(* IEC 61131-3 sources: Antarbhukti-LLM/DatasetCreation/SeedSTs/batch2_filtered_NETWORK, 29 files *)

(* ---- DLOG_FILE_TO_FTP.ST ---- *)
(*@PROPERTIES_EX@
TYPE: POU
LOCALE: 0
IEC_LANGUAGE: ST
PLC_TYPE: independent
PROC_TYPE: independent
GROUP: DATA_LOG
*)
(*@KEY@:DESCRIPTION*)
version 1.1		26. jul. 2011
programmer		ks
tested by		ks

DLOG_FILE_TO_FTP der Baustein kopiert bzw verschiebt die vom DLOG_STORE_FILE_CSV erzeugten Dateien auf einem FTP-Server

(*@KEY@:END_DESCRIPTION*)
FUNCTION_BLOCK DLOG_FILE_TO_FTP

(*Group:parameter*)

VAR_INPUT
	FTP_URL :	oscat_STRING250;
	FTP_ACTIV :	BOOL;
	FILE_DELETE :	BOOL;
	TIMEOUT :	TIME := T#30s;
	RETRY :	INT;
	RETRY_TIME :	TIME := T#30s;
	DNS_IP4 :	DWORD;
	PLC_IP4 :	DWORD;
END_VAR

VAR_OUTPUT
	DONE :	BOOL;
	BUSY :	BOOL;
	ERROR_C :	DWORD;
	ERROR_T :	BYTE;
END_VAR

VAR_IN_OUT
	X :	oscat_DLOG_DATA;
END_VAR

(*Group:lokal*)

VAR
	UCBD :	oscat_UNI_CIRCULAR_BUFFER_DATA;
	UCB :	UNI_CIRCULAR_BUFFER;
	FTP_CLIENT :	FTP_CLIENT;
	WT_1 :	TON;
	ftrig_old :	BOOL;
	filename :	STRING;
	step :	INT;
	ftp_busy :	BOOL;
	ftp_done :	BOOL;
	cnt :	INT;
END_VAR

(*Group:debug*)

VAR
	(*<LOG_MSG :	LOG_MSG;>*)
END_VAR

VAR_EXTERNAL
	(*<LOG_CL :	us_LOG_CONTROL;>*)(*Debug-Datenstruktur*)
END_VAR

VAR
	(*<_debug_enable :	BOOL := TRUE;>*)
END_VAR

(*@KEY@: WORKSHEET
NAME: DLOG_FILE_TO_FTP
IEC_LANGUAGE: ST
*)
(* neue Filenamen speichern *)
IF X.NEW_FILE_RTRIG AND ftrig_old = FALSE THEN
	UCBD.D_HEAD := WORD#1;
	UCBD.D_MODE := 1;
	UCBD.D_STRING := X.NEW_FILE;
	UCB(DATA:=UCBD); (* Daten eintragen *)
	UCBD := UCB.DATA;
END_IF;
ftrig_old := X.NEW_FILE_RTRIG;

CASE step OF

00:	IF UCBD.BUF_COUNT > 0 AND ftp_busy = FALSE THEN
		UCBD.D_MODE := 12; (* Daten lesen und löschen *)
		UCB(DATA:=UCBD);
		UCBD := UCB.DATA;
		filename := UCBD.D_STRING;
		cnt := 0;
		step := 10;
	END_IF;

10:	IF ftp_busy = FALSE THEN
		IF ftp_done THEN
			(*####################  DEBUG-MESSAGE  ###################################*)
			(*IF _debug_enable THEN
				LOG_CL.NEW_MSG := 'F_T_FTP: /FILE OK >~1<';
				LOG_CL.PRINTF[1] := filename;
				LOG_MSG();
			END_IF;*)
			(*########################################################################*)
			step := 0;
		ELSE
			step := 20; (* pause nach error *)
		END_IF;
	END_IF;

20:	IF WT_1.Q THEN (* Wartezeit *)
		cnt := cnt - 1;
		IF RETRY = 0 THEN (* FTP Transfer unbegrenzt wiederholen *)
			(*####################  DEBUG-MESSAGE  ###################################*)
			(*IF _debug_enable THEN
				LOG_CL.NEW_MSG := 'F_T_FTP: Auftrag unbegrenzt wiederholen /file: ~2';
				LOG_CL.PRINTF[2] := filename;
				LOG_MSG();
			END_IF;*)
			(*########################################################################*)
			step := 10; (* FTP Transfer wiederholen *)
		ELSIF cnt >= 0 THEN
			(*####################  DEBUG-MESSAGE  ###################################*)
			(*IF _debug_enable THEN
				LOG_CL.NEW_MSG := 'F_T_FTP: Auftrag wiederholen /cnt: ~1 /file: ~2';
				LOG_CL.PRINTF[1] := INT_TO_STRING(cnt,'%d');
				LOG_CL.PRINTF[2] := filename;
				LOG_MSG();
			END_IF;*)
			(*########################################################################*)
			step := 10; (* FTP Transfer wiederholen *)
		ELSE
			(*####################  DEBUG-MESSAGE  ###################################*)
			(*IF _debug_enable THEN
				LOG_CL.NEW_MSG := 'F_T_FTP: Auftrag verworfen /file: ~2';
				LOG_CL.PRINTF[2] := filename;
				LOG_MSG();
			END_IF;*)
			(*########################################################################*)
			step := 0; (* FTP Auftrag verwerfen *)
		END_IF;
	END_IF;

END_CASE;

BUSY := step = 10;
DONE := step = 0;
WT_1(IN:= step = 20, PT:= RETRY_TIME);

FTP_CLIENT(
	ACTIVATE:= BUSY,
	FILENAME:= filename,
	FTP_URL:= FTP_URL,
	FTP_DOWNLOAD:= FALSE,
	FTP_ACTIV:= FTP_ACTIV,
	FILE_DELETE:= FILE_DELETE,
	TIMEOUT:= TIMEOUT,
	DNS_IP4:= DNS_IP4,
	PLC_IP4:= PLC_IP4
	);
	ftp_done := FTP_CLIENT.DONE;
	ftp_busy := FTP_CLIENT.BUSY;
	ERROR_C := FTP_CLIENT.ERROR_C;
	ERROR_T := FTP_CLIENT.ERROR_T;

(* revision history
ks	01. jan. 2011	rev 1.0
	original version

ks	26. jul. 2011	rev 1.1
    codeoptimierung D_MODE 12

*)

(*@KEY@: END_WORKSHEET *)
END_FUNCTION_BLOCK

(* ---- DLOG_FILE_TO_SMTP.ST ---- *)
(*@PROPERTIES_EX@
TYPE: POU
LOCALE: 0
IEC_LANGUAGE: ST
PLC_TYPE: independent
PROC_TYPE: independent
GROUP: DATA_LOG
*)
(*@KEY@:DESCRIPTION*)
version 1.2		26. jul. 2011
programmer		ks
tested by		ks

DLOG_FILE_TO_SMTP der Baustein versendet die vom DLOG_STORE_FILE_CSV erzeugten Dateien als Email

(*@KEY@:END_DESCRIPTION*)
FUNCTION_BLOCK DLOG_FILE_TO_SMTP

(*Group:parameter*)

VAR_INPUT
	FILE_DELETE :	BOOL;
	TIMEOUT :	TIME := T#30s;
	DTI :	UDINT;
	DTI_OFFSET :	INT;
	RETRY :	INT;
	RETRY_TIME :	TIME := T#30s;
	DNS_IP4 :	DWORD;
END_VAR

VAR_OUTPUT
	DONE :	BOOL;
	BUSY :	BOOL;
	ERROR_C :	DWORD;
	ERROR_T :	BYTE;
END_VAR

VAR_IN_OUT
	SERVER :	STRING;
	MAILFROM :	STRING;
	MAILTO :	oscat_STRING250;
	SUBJECT :	STRING;
	BODY :	oscat_STRING250;
	X :	oscat_DLOG_DATA;
END_VAR

(*Group:lokal*)

VAR
	UCBD :	oscat_UNI_CIRCULAR_BUFFER_DATA;
	UCB :	UNI_CIRCULAR_BUFFER;
	SMTP_CLIENT :	SMTP_CLIENT;
	WT_1 :	TON;
	ftrig_old :	BOOL;
	files :	oscat_STRING250;
	step :	INT;
	smtp_busy :	BOOL;
	smtp_done :	BOOL;
	cnt :	INT;
END_VAR

(*Group:debug*)

VAR
	(*<LOG_MSG :	LOG_MSG;>*)
END_VAR

VAR_EXTERNAL
	(*<LOG_CL :	us_LOG_CONTROL;>*)(*Debug-Datenstruktur*)
END_VAR

VAR
	(*<_debug_enable :	BOOL := TRUE;>*)
END_VAR

(*@KEY@: WORKSHEET
NAME: DLOG_FILE_TO_SMTP
IEC_LANGUAGE: ST
*)
(* neue Filenamen speichern *)
IF X.NEW_FILE_RTRIG AND ftrig_old = FALSE THEN
	UCBD.D_HEAD := WORD#1;
	UCBD.D_MODE := 1;
	UCBD.D_STRING := X.NEW_FILE;
	UCB(DATA:=UCBD); (* Daten eintragen *)
	UCBD := UCB.DATA;
END_IF;
ftrig_old := X.NEW_FILE_RTRIG;

CASE step OF

00:	IF UCBD.BUF_COUNT > 0 AND smtp_busy = FALSE THEN
		UCBD.D_MODE := 12; (* Daten lesen und löschen *)
		UCB(DATA:=UCBD);
		UCBD := UCB.DATA;
		files := UCBD.D_STRING;
		IF FILE_DELETE THEN
			files := CONCAT(files,';#DEL#');
		END_IF;
		cnt := 0;
		step := 10;
	END_IF;

10:	IF smtp_busy = FALSE THEN
		IF smtp_done THEN
			(*####################  DEBUG-MESSAGE  ###################################*)
			(*IF _debug_enable THEN
				LOG_CL.NEW_MSG := 'F_T_SMTP: /FILE OK >~1<';
				LOG_CL.PRINTF[1] := files;
				LOG_MSG();
			END_IF;*)
			(*########################################################################*)
			step := 0;
		ELSE
			step := 20; (* pause nach error *)
		END_IF;
	END_IF;

20:	IF WT_1.Q THEN (* Wartezeit *)
		cnt := cnt - 1;
		IF RETRY = 0 THEN (* Transfer unbegrenzt wiederholen *)
			(*####################  DEBUG-MESSAGE  ###################################*)
			(*IF _debug_enable THEN
				LOG_CL.NEW_MSG := 'F_T_SMTP: Auftrag unbegrenzt wiederholen /file: ~2';
				LOG_CL.PRINTF[2] := files;
				LOG_MSG();
			END_IF;*)
			(*########################################################################*)
			step := 10; (* Transfer wiederholen *)
		ELSIF cnt >= 0 THEN
			(*####################  DEBUG-MESSAGE  ###################################*)
			(*IF _debug_enable THEN
				LOG_CL.NEW_MSG := 'F_T_SMTP: Auftrag wiederholen /cnt: ~1 /file: ~2';
				LOG_CL.PRINTF[1] := INT_TO_STRING(cnt,'%d');
				LOG_CL.PRINTF[2] := files;
				LOG_MSG();
			END_IF;*)
			(*########################################################################*)
			step := 10; (* Transfer wiederholen *)
		ELSE
			(*####################  DEBUG-MESSAGE  ###################################*)
			(*IF _debug_enable THEN
				LOG_CL.NEW_MSG := 'F_T_SMTP: Auftrag verworfen /file: ~2';
				LOG_CL.PRINTF[2] := files;
				LOG_MSG();
			END_IF;*)
			(*########################################################################*)
			step := 0; (* Auftrag verwerfen *)
		END_IF;
	END_IF;

END_CASE;

BUSY := step = 10;
DONE := step = 0;
WT_1(IN:= step = 20, PT:= RETRY_TIME);

SMTP_CLIENT(
	ACTIVATE:= BUSY,
	TIMEOUT:= TIMEOUT,
	DTI:= DTI,
	DTI_OFFSET:= DTI_OFFSET,
	DNS_IP4:= DNS_IP4,
	SERVER:= SERVER,
	MAILFROM:= MAILFROM,
	MAILTO:= MAILTO,
	SUBJECT:= SUBJECT,
	BODY:= BODY,
	FILES:= FILES
	);
	SERVER:= SMTP_CLIENT.SERVER;
	MAILFROM:= SMTP_CLIENT.MAILFROM;
	MAILTO:= SMTP_CLIENT.MAILTO;
	SUBJECT:= SMTP_CLIENT.SUBJECT;
	BODY:= SMTP_CLIENT.BODY;
	FILES:= SMTP_CLIENT.FILES;
	smtp_done := SMTP_CLIENT.DONE;
	smtp_busy := SMTP_CLIENT.BUSY;
	ERROR_C := SMTP_CLIENT.ERROR_C;
	ERROR_T := SMTP_CLIENT.ERROR_T;

(* revision history

ks	01. jan. 2011	rev 1.0
	original version

ks	28. apr. 2011	rev 1.1
	stringfehler bei option 'file_delete'

ks	26. jul. 2011	rev 1.2
    codeoptimierung D_MODE 12
*)

(*@KEY@: END_WORKSHEET *)
END_FUNCTION_BLOCK

(* ---- DLOG_STORE_FILE_CSV.ST ---- *)
(*@PROPERTIES_EX@
TYPE: POU
LOCALE: 0
IEC_LANGUAGE: ST
PLC_TYPE: independent
PROC_TYPE: independent
GROUP: DATA_LOG
*)
(*@KEY@:DESCRIPTION*)
version 1.2		25. jul. 2011
programmer		ks
tested by		ks

DLOG_STORE_FILE_CSV der Baustein schreibt die DLOG Parameter in einen lokale Datei im CSV-Format

(*@KEY@:END_DESCRIPTION*)
FUNCTION_BLOCK DLOG_STORE_FILE_CSV

(*Group:Default*)

VAR_INPUT
	ENABLE :	BOOL;
	TRIG_M :	BOOL;
	TRIG_T :	UDINT;
	FILENAME :	STRING;
	DTI :	UDINT;
	SEP :	BYTE;
END_VAR

VAR_OUTPUT
	ERROR_C :	DWORD;
	ERROR_T :	BYTE;
END_VAR

VAR_IN_OUT
	X :	oscat_DLOG_DATA;
END_VAR

VAR
	FS :	FILE_SERVER;
	FSD :	oscat_FILE_SERVER_DATA;
	PT :	oscat_NETWORK_BUFFER;
	UCB :	UNI_CIRCULAR_BUFFER;
	ra :	BOOL;
	trig_m_last :	BOOL;
	dti_last :	UDINT := udint#4294967295;(*DT#2070-02-06-06:28:15*)
	enable_last :	BOOL;
	fn_last :	STRING;
	fn :	STRING;
	init :	BOOL;
	step :	INT;
	idx :	INT;
	log_stop :	BOOL;
	buf_totalsize :	INT := 4096;
	DT_TO_STRF :	DT_TO_STRF;
	_STRING_TO_BUFFER :	_STRING_TO_BUFFER_NW;
	n :	USINT;
END_VAR

(*@KEY@: WORKSHEET
NAME: DLOG_STORE_FILE_CSV
IEC_LANGUAGE: ST
*)
X.DTI := DTI; (* Datum / Zeit eintragen *)
IF DTI <> dti_last THEN
	X.CLOCK_TRIG := TRUE;
	dti_last := DTI;
	X.STORE_TYPE := BYTE#2;
ELSE
	X.CLOCK_TRIG := FALSE;
END_IF;

IF X.ADD_HEADER = FALSE THEN (* wenn add-header und add-data gleichzeitig ansteht, dann add-data einen zyklus länger anstehen lassen *)
	X.ADD_DATA := FALSE;
END_IF;
X.ADD_HEADER := FALSE;

IF ENABLE THEN
	IF X.CLOCK_TRIG THEN
		DT_TO_STRF(DTI:=DTI,MS:=0,FMT:=FILENAME,LANG:=0); (* automatische Dateinamen generierung *)
		fn := DT_TO_STRF.DT_TO_STRF;
		IF TRIG_T > UDINT#0 THEN (* automatischer Trigger *)
			ra := DTI MOD TRIG_T = UDINT#0;
		END_IF;
	ELSE
		ra := FALSE;
	END_IF;
	IF (TRIG_M AND NOT trig_m_last) OR ra THEN (* manueller oder automatischer Trigger *)
		X.ADD_DATA := TRUE; (* Daten loggen *)
	END_IF;
	IF NOT init THEN
		init := TRUE;
		X.ADD_HEADER := TRUE; (* Spaltenüberschriften übernehmen *)
	END_IF;
END_IF;

IF (NOT ENABLE AND enable_last) OR (NE_STRING(fn,fn_last) AND step > 0) THEN (* Neg. Flanke ENABLE - Log Stop *)
	fn_last := fn;
	X.UCB.D_HEAD := WORD#16#FF00;
	X.UCB.D_MODE := 1;
	UCB(DATA:=X.UCB); (* Element schreiben *)
	X.UCB := UCB.DATA;
	X.ADD_HEADER := TRUE; (* Spaltenüberschriften übernehmen *)
END_IF;

CASE step OF

00:	IF ENABLE THEN
		fn_last := fn;
		FSD.FILENAME := fn; (* Dateiname *)
		FSD.OFFSET := UDINT#0; (* Start bei Dateianfang *)
		FSD.AUTO_CLOSE := T#0s; (* Auto-Close *)
		step := 20;
	END_IF;

20:	IF X.UCB.BUF_COUNT > 0 THEN (* Einträge vorhanden *)
		X.UCB.D_MODE := 10;
		UCB(DATA:=X.UCB); (* Element lesen , aber noch nicht entfernen *)
		X.UCB := UCB.DATA;
		IF X.UCB.D_HEAD = WORD#16#FF00 THEN (* LOG_STOP Command *)
			X.UCB.D_MODE := 11;
			UCB(DATA:=X.UCB); (* Element entfernen *)
			X.UCB := UCB.DATA;
			log_stop := TRUE;
			step := 40; (* Daten schreiben *)
		ELSIF idx + LEN(X.UCB.D_STRING) + 2 < buf_totalsize THEN (* Platz für Element vorhanden ? *)
			X.UCB.D_MODE := 11;
			UCB(DATA:=X.UCB); (* Element entfernen *)
			X.UCB := UCB.DATA;
			_STRING_TO_BUFFER(STR:=X.UCB.D_STRING, POS:=idx, PT:=PT.BUFFER, SIZE:=INT_TO_UINT(buf_totalsize));
			PT.BUFFER:=_STRING_TO_BUFFER.PT;
			idx := idx + LEN(X.UCB.D_STRING);
			n := n + USINT#1;
			IF n = X.ID_MAX THEN (* letztes Element einer Zeile *)
				n := USINT#0;
				PT.BUFFER[idx] := BYTE#16#0D;
				idx := idx + 1;
				PT.BUFFER[idx] := BYTE#16#0A;
			ELSE
				PT.BUFFER[idx] := SEP;
			END_IF;
			idx := idx + 1;
		ELSE
			step := 40; (* Daten schreiben *)
		END_IF;
	END_IF;

40:	IF idx > 0 THEN (* Daten schreiben *)
		FSD.MODE := BYTE#3; (* create + write *)
		PT.SIZE := INT_TO_UINT(idx); (* Datenlänge eintragen *)
		idx := 0;
	END_IF;
	step := 60;

60:	IF FSD.MODE = BYTE#0 THEN
		IF log_stop THEN
			log_stop := FALSE;
			FSD.MODE := BYTE#5; (* Datei schliessen *)
			X.NEW_FILE := FSD.FILENAME;
			X.NEW_FILE_RTRIG := FALSE;
			step := 80;
		ELSE
			step := 20;
		END_IF;
	END_IF;

80:	IF FSD.MODE = BYTE#0 THEN (* Datei schliessen beendet *)
		X.NEW_FILE_RTRIG := TRUE;
		step := 0;
	END_IF;

END_CASE;

trig_m_last := TRIG_M;
enable_last := ENABLE;

FS(FSD:=FSD,PT:=PT); (* FILE_SERVER *)
FSD := FS.FSD;
PT  := FS.PT;

ERROR_C := BYTE_TO_DWORD(FSD.ERROR);
ERROR_T := SEL(FSD.ERROR > BYTE#0,BYTE#0,BYTE#1);

(* revision history
ks	01. jan. 2011	rev 1.0
	original version

ks	13. may. 2011	rev 1.1
	ADD_DATA_REQ, ERROR_T, ERROR_C hinzugefügt

ks	25. jul. 2011	rev 1.2
	HEAD informationen geändert, neuer Spaltenzähler

*)

(*@KEY@: END_WORKSHEET *)
END_FUNCTION_BLOCK

(* ---- DLOG_STORE_FILE_HTML.ST ---- *)
(*@PROPERTIES_EX@
TYPE: POU
LOCALE: 0
IEC_LANGUAGE: ST
PLC_TYPE: independent
PROC_TYPE: independent
GROUP: DATA_LOG
*)
(*@KEY@:DESCRIPTION*)

(*@KEY@:END_DESCRIPTION*)
FUNCTION_BLOCK DLOG_STORE_FILE_HTML

(*Group:Default*)

VAR_INPUT
	ENABLE :	BOOL;
	TRIG_M :	BOOL;
	TRIG_T :	UDINT;
	FILENAME :	STRING;
	DTI :	UDINT;
	HTML_CAPTION :	STRING;
	HTML_TABLE :	STRING;
	HTML_TR_HEAD :	STRING;
	HTML_TR_EVEN :	STRING;
	HTML_TR_ODD :	STRING;
END_VAR

VAR_OUTPUT
	ERROR_C :	DWORD;
	ERROR_T :	BYTE;
END_VAR

VAR_IN_OUT
	X :	oscat_DLOG_DATA;
END_VAR

VAR
	FS :	FILE_SERVER;
	FSD :	oscat_FILE_SERVER_DATA;
	PT :	oscat_NETWORK_BUFFER;
	UCB :	UNI_CIRCULAR_BUFFER;
	ra :	BOOL;
	trig_m_last :	BOOL;
	dti_last :	UDINT := udint#4294967295;(*DT#2070-02-06-06:28:15*)
	enable_last :	BOOL;
	fn_last :	STRING;
	str :	oscat_STRING250;
	fn :	STRING;
	init :	BOOL;
	step :	INT;
	idx :	INT;
	log_state :	USINT;
	color :	BOOL;
	head :	BOOL;
	n :	USINT;
	buf_totalsize :	INT := 4096;
	DT_TO_STRF :	DT_TO_STRF;
	_STRING_TO_BUFFER :	_STRING_TO_BUFFER_NW;
END_VAR

(*@KEY@: WORKSHEET
NAME: DLOG_STORE_FILE_HTML
IEC_LANGUAGE: ST
*)
X.DTI := DTI; (* Datum / Zeit eintragen *)
IF DTI <> dti_last THEN
	X.CLOCK_TRIG := TRUE;
	dti_last := DTI;
	X.STORE_TYPE := BYTE#4;
ELSE
	X.CLOCK_TRIG := FALSE;
END_IF;

IF X.ADD_HEADER = FALSE THEN (* wenn add-header und add-data gleichzeitig ansteht, dann add-data einen zyklus länger anstehen lassen *)
	X.ADD_DATA := FALSE;
END_IF;
X.ADD_HEADER := FALSE;

IF ENABLE THEN
	IF X.CLOCK_TRIG THEN
		DT_TO_STRF(DTI:=DTI,MS:=0,FMT:=FILENAME,LANG:=0); (* automatische Dateinamen generierung *)
		fn := DT_TO_STRF.DT_TO_STRF;
		IF TRIG_T > UDINT#0 THEN (* automatischer Trigger *)
			ra := DTI MOD TRIG_T = UDINT#0;
		END_IF;
	ELSE
		ra := FALSE;
	END_IF;
	IF (TRIG_M AND NOT trig_m_last) OR ra OR X.ADD_DATA_REQ THEN (* manueller, automatischer oder externer Trigger *)
		X.ADD_DATA := TRUE; (* Daten loggen *)
	END_IF;
	IF NOT init THEN
		init := TRUE;
		X.ADD_HEADER := TRUE; (* Spaltenüberschriften übernehmen *)
	END_IF;
END_IF;
X.ADD_DATA_REQ := FALSE; (* externe Anforderung rücksetzen *)

IF (NOT ENABLE AND enable_last) OR (NE_STRING(fn,fn_last) AND step > 0) THEN (* Neg. Flanke ENABLE - Log Stop *)
	fn_last := fn;
	X.UCB.D_HEAD := WORD#16#FF00;
	X.UCB.D_MODE := 1;
	UCB(DATA:=X.UCB); (* Element schreiben *)
	X.UCB := UCB.DATA;
	X.ADD_HEADER := TRUE; (* Spaltenüberschriften übernehmen *)
END_IF;

CASE step OF

00:	IF ENABLE THEN
		color := FALSE;
		head := FALSE;
		fn_last := fn;
		FSD.FILENAME := fn; (* Dateiname *)
		FSD.OFFSET := UDINT#0; (* Start bei Dateianfang *)
		FSD.AUTO_CLOSE := T#0s; (* Auto-Close *)
		step := 10;
	END_IF;

10:	(* Headerdaten schreiben *)
	str := CONCAT('<html><body><table ',HTML_TABLE);
	str := CONCAT(str,'><caption>');
	str := CONCAT(str,HTML_CAPTION);
	str := CONCAT(str,'</caption>');

	_STRING_TO_BUFFER(STR:=str, POS:=idx, PT:=PT.BUFFER, SIZE:=INT_TO_UINT(buf_totalsize));
	PT.BUFFER:=_STRING_TO_BUFFER.PT;
	idx := idx + LEN(str);
	step := 20;

20:	IF log_state = USINT#254 THEN
		log_state := USINT#255;
		str := '</table></body></html>';
		_STRING_TO_BUFFER(STR:=str, POS:=idx, PT:=PT.BUFFER, SIZE:=INT_TO_UINT(buf_totalsize));
		PT.BUFFER:=_STRING_TO_BUFFER.PT;
		idx := idx + LEN(str);
		step := 40; (* Daten schreiben *)

	ELSIF X.UCB.BUF_COUNT > 0 THEN (* Einträge vorhanden *)
		X.UCB.D_MODE := 10;
		UCB(DATA:=X.UCB); (* Element lesen , aber noch nicht entfernen *)
		X.UCB := UCB.DATA;

		IF X.UCB.D_HEAD = WORD#16#FF00 THEN (* LOG_STOP Command *)
			X.UCB.D_MODE := 11;
			UCB(DATA:=X.UCB); (* Element entfernen *)
			X.UCB := UCB.DATA;
			log_state := USINT#254;

		ELSIF idx + LEN(X.UCB.D_STRING) + 120 < buf_totalsize THEN (* Platz für Element vorhanden ? *)
			X.UCB.D_MODE := 11;
			UCB(DATA:=X.UCB); (* Element entfernen *)
			X.UCB := UCB.DATA;

			IF log_state = USINT#0 THEN
				str := '<TR ';
				IF NOT head THEN
					str := CONCAT(str,HTML_TR_HEAD);
					head := TRUE;
				ELSIF color THEN
					str := CONCAT(str,HTML_TR_EVEN);
				ELSE
					str := CONCAT(str,HTML_TR_ODD);
				END_IF;
				str := CONCAT(str,'><TD>');
			ELSE
				str := '<TD>';
			END_IF;
			_STRING_TO_BUFFER(STR:=str, POS:=idx, PT:=PT.BUFFER, SIZE:=INT_TO_UINT(buf_totalsize));
			PT.BUFFER:=_STRING_TO_BUFFER.PT;
			idx := idx + LEN(str);
			log_state := log_state + USINT#1;

			_STRING_TO_BUFFER(STR:=X.UCB.D_STRING, POS:=idx, PT:=PT.BUFFER, SIZE:=INT_TO_UINT(buf_totalsize));
			PT.BUFFER:=_STRING_TO_BUFFER.PT;
			idx := idx + LEN(X.UCB.D_STRING);
			n := n + USINT#1;
			IF n = X.ID_MAX THEN
				n := USINT#0;
				str := '</TD></TR>';
				color := NOT color;
				log_state := USINT#0;
			ELSE
				str := '</TD>';
			END_IF;
			_STRING_TO_BUFFER(STR:=str, POS:=idx, PT:=PT.BUFFER, SIZE:=INT_TO_UINT(buf_totalsize));
			PT.BUFFER:=_STRING_TO_BUFFER.PT;
			idx := idx + LEN(str);
		END_IF;
		step := 40; (* Daten schreiben *)
	END_IF;

40:	IF idx > 0 THEN (* Daten schreiben *)
		FSD.MODE := BYTE#3; (* create + write *)
		PT.SIZE := INT_TO_UINT(idx); (* Datenlänge eintragen *)
		idx := 0;
	END_IF;
	step := 60;

60:	IF FSD.MODE = BYTE#0 THEN
		IF log_state = USINT#255 THEN
			log_state := USINT#0;
			FSD.MODE := BYTE#5; (* Datei schliessen *)
			X.NEW_FILE := FSD.FILENAME;
			X.NEW_FILE_RTRIG := FALSE;
			step := 80;
		ELSE
			step := 20;
		END_IF;
	END_IF;

80:	IF FSD.MODE = BYTE#0 THEN (* Datei schliessen beendet *)
		X.NEW_FILE_RTRIG := TRUE;
		step := 0;
	END_IF;

END_CASE;

trig_m_last := TRIG_M;
enable_last := ENABLE;

FS(FSD:=FSD,PT:=PT); (* FILE_SERVER *)
FSD := FS.FSD;
PT  := FS.PT;

ERROR_C := BYTE_TO_DWORD(FSD.ERROR);
ERROR_T := SEL(FSD.ERROR > BYTE#0,BYTE#0,BYTE#1);

(* revision history
ks	25. july. 2011	rev 1.0
	original version

*)

(*@KEY@: END_WORKSHEET *)
END_FUNCTION_BLOCK

(* ---- DLOG_STORE_FILE_XML.ST ---- *)
(*@PROPERTIES_EX@
TYPE: POU
LOCALE: 0
IEC_LANGUAGE: ST
PLC_TYPE: independent
PROC_TYPE: independent
GROUP: DATA_LOG
*)
(*@KEY@:DESCRIPTION*)
version 1.0		25. july. 2011
programmer		ks
tested by		ks

DLOG_STORE_FILE_XML schreibt die DLOG Parameter in einen lokale Datei im XML-Format

(*@KEY@:END_DESCRIPTION*)
FUNCTION_BLOCK DLOG_STORE_FILE_XML

(*Group:Default*)

VAR_INPUT
	ENABLE :	BOOL;
	TRIG_M :	BOOL;
	TRIG_T :	UDINT;
	FILENAME :	STRING;
	DTI :	UDINT;
END_VAR

VAR_OUTPUT
	ERROR_C :	DWORD;
	ERROR_T :	BYTE;
END_VAR

VAR_IN_OUT
	X :	oscat_DLOG_DATA;
END_VAR

VAR
	FS :	FILE_SERVER;
	FSD :	oscat_FILE_SERVER_DATA;
	PT :	oscat_NETWORK_BUFFER;
	UCB :	UNI_CIRCULAR_BUFFER;
	ra :	BOOL;
	trig_m_last :	BOOL;
	dti_last :	UDINT := udint#4294967295;(*DT#2070-02-06-06:28:15*)
	enable_last :	BOOL;
	fn_last :	STRING;
	str :	oscat_STRING250;
	fn :	STRING;
	init :	BOOL;
	step :	INT;
	idx :	INT;
	log_state :	USINT;
	n :	USINT;
	buf_totalsize :	INT := 4096;
	DT_TO_STRF :	DT_TO_STRF;
	_STRING_TO_BUFFER :	_STRING_TO_BUFFER_NW;
END_VAR

(*@KEY@: WORKSHEET
NAME: DLOG_STORE_FILE_XML
IEC_LANGUAGE: ST
*)
X.DTI := DTI; (* Datum / Zeit eintragen *)
IF DTI <> dti_last THEN
	X.CLOCK_TRIG := TRUE;
	dti_last := DTI;
	X.STORE_TYPE := BYTE#3;
ELSE
	X.CLOCK_TRIG := FALSE;
END_IF;

IF X.ADD_HEADER = FALSE THEN (* wenn add-header und add-data gleichzeitig ansteht, dann add-data einen zyklus länger anstehen lassen *)
	X.ADD_DATA := FALSE;
END_IF;
X.ADD_HEADER := FALSE;

IF ENABLE THEN
	IF X.CLOCK_TRIG THEN
		DT_TO_STRF(DTI:=DTI,MS:=0,FMT:=FILENAME,LANG:=0); (* automatische Dateinamen generierung *)
		fn := DT_TO_STRF.DT_TO_STRF;
		IF TRIG_T > UDINT#0 THEN (* automatischer Trigger *)
			ra := DTI MOD TRIG_T = UDINT#0;
		END_IF;
	ELSE
		ra := FALSE;
	END_IF;
	IF (TRIG_M AND NOT trig_m_last) OR ra OR X.ADD_DATA_REQ THEN (* manueller, automatischer oder externer Trigger *)
		X.ADD_DATA := TRUE; (* Daten loggen *)
	END_IF;
	IF NOT init THEN
		init := TRUE;
		X.ADD_HEADER := TRUE; (* Spaltenüberschriften übernehmen *)
	END_IF;
END_IF;
X.ADD_DATA_REQ := FALSE; (* externe Anforderung rücksetzen *)

IF (NOT ENABLE AND enable_last) OR (NE_STRING(fn,fn_last) AND step > 0) THEN (* Neg. Flanke ENABLE - Log Stop *)
	fn_last := fn;
	X.UCB.D_HEAD := WORD#16#FF00;
	X.UCB.D_MODE := 1;
	UCB(DATA:=X.UCB); (* Element schreiben *)
	X.UCB := UCB.DATA;
	X.ADD_HEADER := TRUE; (* Spaltenüberschriften übernehmen *)
END_IF;

CASE step OF

00:	IF ENABLE THEN
		fn_last := fn;
		FSD.FILENAME := fn; (* Dateiname *)
		FSD.OFFSET := UDINT#0; (* Start bei Dateianfang *)
		FSD.AUTO_CLOSE := T#0s; (* Auto-Close *)
		step := 10;
	END_IF;

10:	(* Headerdaten schreiben *)
	str := '<?xml version="1.0" encoding="UTF-8"?><table>';
	_STRING_TO_BUFFER(STR:=str, POS:=idx, PT:=PT.BUFFER, SIZE:=INT_TO_UINT(buf_totalsize));
	PT.BUFFER:=_STRING_TO_BUFFER.PT;
	idx := idx + LEN(str);
	step := 20;

20:	IF log_state = USINT#254 THEN
		log_state := USINT#255;
		str := '</table>';
		_STRING_TO_BUFFER(STR:=str, POS:=idx, PT:=PT.BUFFER, SIZE:=INT_TO_UINT(buf_totalsize));
		PT.BUFFER:=_STRING_TO_BUFFER.PT;
		idx := idx + LEN(str);
		step := 40; (* Daten schreiben *)

	ELSIF X.UCB.BUF_COUNT > 0 THEN (* Einträge vorhanden *)
		X.UCB.D_MODE := 10;
		UCB(DATA:=X.UCB); (* Element lesen , aber noch nicht entfernen *)
		X.UCB := UCB.DATA;

		IF X.UCB.D_HEAD = WORD#16#FF00 THEN (* LOG_STOP Command *)
			X.UCB.D_MODE := 11;
			UCB(DATA:=X.UCB); (* Element entfernen *)
			X.UCB := UCB.DATA;
			log_state := USINT#254;

		ELSIF idx + LEN(X.UCB.D_STRING) + 120 < buf_totalsize THEN (* Platz für Element vorhanden ? *)
			X.UCB.D_MODE := 11;
			UCB(DATA:=X.UCB); (* Element entfernen *)
			X.UCB := UCB.DATA;

			IF log_state = USINT#0 THEN
				str := '<row><entry>';
			ELSE
				str := '<entry>';
			END_IF;

			_STRING_TO_BUFFER(STR:=str, POS:=idx, PT:=PT.BUFFER, SIZE:=INT_TO_UINT(buf_totalsize));
			PT.BUFFER:=_STRING_TO_BUFFER.PT;
			idx := idx + LEN(str);
			log_state := log_state + USINT#1;

			_STRING_TO_BUFFER(STR:=X.UCB.D_STRING, POS:=idx, PT:=PT.BUFFER, SIZE:=INT_TO_UINT(buf_totalsize));
			PT.BUFFER:=_STRING_TO_BUFFER.PT;
			idx := idx + LEN(X.UCB.D_STRING);

			n := n + USINT#1;
			IF n = X.ID_MAX THEN
				n := USINT#0;
				str := '</entry></row>';
				log_state := USINT#0;
			ELSE
				str := '</entry>';
			END_IF;
			_STRING_TO_BUFFER(STR:=str, POS:=idx, PT:=PT.BUFFER, SIZE:=INT_TO_UINT(buf_totalsize));
			PT.BUFFER:=_STRING_TO_BUFFER.PT;
			idx := idx + LEN(str);
		END_IF;
		step := 40; (* Daten schreiben *)
	END_IF;

40:	IF idx > 0 THEN (* Daten schreiben *)
		FSD.MODE := BYTE#3; (* create + write *)
		PT.SIZE := INT_TO_UINT(idx); (* Datenlänge eintragen *)
		idx := 0;
	END_IF;
	step := 60;

60:	IF FSD.MODE = BYTE#0 THEN
		IF log_state = USINT#255 THEN
			log_state := USINT#0;
			FSD.MODE := BYTE#5; (* Datei schliessen *)
			X.NEW_FILE := FSD.FILENAME;
			X.NEW_FILE_RTRIG := FALSE;
			step := 80;
		ELSE
			step := 20;
		END_IF;
	END_IF;

80:	IF FSD.MODE = BYTE#0 THEN (* Datei schliessen beendet *)
		X.NEW_FILE_RTRIG := TRUE;
		step := 0;
	END_IF;

END_CASE;

trig_m_last := TRIG_M;
enable_last := ENABLE;

FS(FSD:=FSD,PT:=PT); (* FILE_SERVER *)
FSD := FS.FSD;
PT  := FS.PT;

ERROR_C := BYTE_TO_DWORD(FSD.ERROR);
ERROR_T := SEL(FSD.ERROR > BYTE#0,BYTE#0,BYTE#1);

(* revision history
ks	25. july. 2011	rev 1.0
	original version

*)
(*@KEY@: END_WORKSHEET *)
END_FUNCTION_BLOCK

(* ---- DLOG_STORE_RRD.ST ---- *)
(*@PROPERTIES_EX@
TYPE: POU
LOCALE: 0
IEC_LANGUAGE: ST
PLC_TYPE: independent
PROC_TYPE: independent
GROUP: DATA_LOG
*)
(*@KEY@:DESCRIPTION*)
version 1.2		26. jul. 2011
programmer		ks
tested by		ks

DLOG_STORE_RRD der Baustein übergibt die DLOG Parameter an einen RoundRobinDatabase-Server

(*@KEY@:END_DESCRIPTION*)
FUNCTION_BLOCK DLOG_STORE_RRD

(*Group:Default*)

VAR_INPUT
	ENABLE :	BOOL;
	TRIG_M :	BOOL;
	TRIG_T :	UDINT;
	URL :	oscat_STRING250;
	DTI :	UDINT;
	SEP :	BYTE;
	DNS_IP4 :	DWORD;
	TIMEOUT :	TIME;
END_VAR

VAR_OUTPUT
	ERROR_C :	DWORD;
	ERROR_T :	BYTE;
END_VAR

VAR_IN_OUT
	X :	oscat_DLOG_DATA;
END_VAR

VAR
	UCB :	UNI_CIRCULAR_BUFFER;
	IP_C :	oscat_IP_C;
	S_BUF :	oscat_NETWORK_BUFFER;
	R_BUF :	oscat_NETWORK_BUFFER;
	URL_DATA :	oscat_url;
	DNS_CLIENT :	DNS_CLIENT;
	HTTP_GET :	HTTP_GET;
	IPC :	IP_CONTROL;
	ra :	BOOL;
	trig_m_last :	BOOL;
	dti_last :	UDINT := udint#4294967295;(*DT#2070-02-06-06:28:15*)
	step :	INT;
	sep_char :	oscat_STRING1;
	STRING_TO_URL :	STRING_TO_URL;
	CHR_TO_STRING :	CHR_TO_STRING;
	n :	INT;
END_VAR

(*@KEY@: WORKSHEET
NAME: DLOG_STORE_RRD
IEC_LANGUAGE: ST
*)
X.DTI := DTI; (* Datum / Zeit eintragen *)
IF DTI <> dti_last THEN
	X.CLOCK_TRIG := TRUE;
	dti_last := DTI;
	X.STORE_TYPE := BYTE#1;
ELSE
	X.CLOCK_TRIG := FALSE;
END_IF;

X.ADD_DATA := FALSE;

IF ENABLE THEN
	IF X.CLOCK_TRIG THEN
		IF TRIG_T > UDINT#0 THEN (* automatischer Trigger *)
			ra := DTI MOD TRIG_T = UDINT#0;
		END_IF;
	ELSE
		ra := FALSE;
	END_IF;
	IF (TRIG_M AND NOT trig_m_last) OR ra OR X.ADD_DATA_REQ THEN (* manueller, automatischer oder externer Trigger *)
		X.ADD_DATA := TRUE; (* Daten loggen *)
	END_IF;
END_IF;
X.ADD_DATA_REQ := FALSE; (* externe Anforderung rücksetzen *)

CASE step OF

00:	IF ENABLE THEN
		STRING_TO_URL(STR:=URL,DEFAULT_PROTOCOL:='',DEFAULT_PATH:=''); (* URL zerlegen *)
		URL_DATA:=STRING_TO_URL.STRING_TO_URL;
		CHR_TO_STRING(C:=SEP);
		sep_char:=CHR_TO_STRING.CHR_TO_STRING;
		ERROR_T := BYTE#0;
		ERROR_C := DWORD#0;
		step := 20;
	END_IF;

20:	IF X.UCB.BUF_COUNT >= USINT_TO_INT(X.ID_MAX) THEN (* Einträge vorhanden *)
		n := 1;
		WHILE n <= USINT_TO_INT(X.ID_MAX) DO
			X.UCB.D_MODE := 12; (* Element lesen und löschen *)
			UCB(DATA:=X.UCB);
			X.UCB := UCB.DATA;
			IF n < USINT_TO_INT(X.ID_MAX) THEN (* Trennzeichen hinzufügen *)
				X.UCB.D_STRING := CONCAT(X.UCB.D_STRING,sep_char);
			END_IF;
			IF LEN(X.UCB.D_STRING) + LEN(URL_DATA.QUERY) <= 250 THEN
				URL_DATA.QUERY := CONCAT(URL_DATA.QUERY,X.UCB.D_STRING); (* Query mit LOG-Daten ergänzen *)
				step :=40;
			ELSE
				ERROR_T := BYTE#4; (* LOG-Daten können nicht in URL gepackt werden *)
				ERROR_C := DWORD#1;
				step := 0;
			END_IF;
			n := n + 1;
		END_WHILE;;
	END_IF;

40:	IF DNS_CLIENT.DONE THEN
		step := 60;
	ELSIF (DNS_CLIENT.ERROR > DWORD#0) THEN
		ERROR_C := DNS_CLIENT.ERROR; (* Fehlerbehandlung *)
		ERROR_T := BYTE#1;
		step := 100;
	END_IF;

60:	IF HTTP_GET.DONE THEN
		n := UINT_TO_INT(HTTP_GET.BODY_START);
		IF R_BUF.BUFFER[n] <> BYTE#48 THEN (* ASCII '0' *)
			ERROR_C := DWORD#1;
			ERROR_T := BYTE#3;
		END_IF;
		step := 100;

	ELSIF HTTP_GET.ERROR > DWORD#0 THEN (* Fehlerbehandlung *)
		ERROR_C := HTTP_GET.ERROR;
		ERROR_T := BYTE#2;
		step := 100;
	END_IF;

100:	IF (NOT HTTP_GET.DONE) THEN (* UNLOCK HTTP DATA *)
		step := SEL(ERROR_T = BYTE#0, 120,0);
	END_IF;

120:	IF NOT ENABLE THEN
		X.UCB.D_MODE := 99;
		UCB(DATA:=X.UCB); (* Buffer löschen *)
		X.UCB := UCB.DATA;
		step := 0;
	END_IF;

END_CASE;

HTTP_GET(IP_C:=IP_C,S_BUF:=S_BUF,R_BUF:=R_BUF,IP4:=DNS_CLIENT.IP4,GET:=step=60,MODE:=BYTE#2,UNLOCK_BUF:=step=100,URL_DATA:=URL_DATA); (* HTTP_GET *)
IP_C     := HTTP_GET.IP_C;
S_BUF    := HTTP_GET.S_BUF;
R_BUF    := HTTP_GET.R_BUF;
URL_DATA := HTTP_GET.URL_DATA;

DNS_CLIENT(IP_C:=IP_C, S_BUF:=S_BUF, R_BUF:=R_BUF, DOMAIN:=URL_DATA.DOMAIN, IP4_DNS:= DNS_IP4, ACTIVATE:=step=40); (* DNS-Client *)
IP_C  := DNS_CLIENT.IP_C;
S_BUF := DNS_CLIENT.S_BUF;
R_BUF := DNS_CLIENT.R_BUF;

IPC(IP:= DWORD#0, PORT:= WORD#0 , TIME_OUT:= TIMEOUT, IP_C:= IP_C, S_BUF:= S_BUF, R_BUF:= R_BUF); (* IP_CONTROL *)
IP_C  := IPC.IP_C;
S_BUF := IPC.S_BUF;
R_BUF := IPC.R_BUF;

trig_m_last := TRIG_M;

(* revision history
ks	01. jan. 2011	rev 1.0
	original version

ks	13. may. 2011	rev 1.1
	ADD_DATA_REQ hinzugefügt

ks	26. july. 2011	rev 1.2
	code optimierung D_MODE 12 und bessere fehlerauswertung
*)

(*@KEY@: END_WORKSHEET *)
END_FUNCTION_BLOCK

(* ---- DNS_CLIENT.ST ---- *)
(*@PROPERTIES_EX@
TYPE: POU
LOCALE: 0
IEC_LANGUAGE: ST
PLC_TYPE: independent
PROC_TYPE: independent
GROUP: NETWORK
*)
(*@KEY@:DESCRIPTION*)

version 1.3		26. jul. 2011
programmer 		ks
tested by		ks

DNS_CLIENT führt eine Domain-Name Abfrage bei einen DNS-Server durch
(*@KEY@:END_DESCRIPTION*)
FUNCTION_BLOCK DNS_CLIENT

(*Group:log*)

VAR
	(*<LOG_MSG :	LOG_MSG;>*)
	(*<_debug_enable :	BOOL := FALSE;>*)
END_VAR

VAR_EXTERNAL
	(*<LOG_CL :	us_LOG_CONTROL;>*)
END_VAR

(*Group:lokal*)

VAR
	IP4_DECODE :	IP4_DECODE;
	IP_FIFO :	IP_FIFO;
	CODE :	CODE;
	ip_state :	BYTE;
	ip_id :	BYTE;
	i :	INT;
	i1 :	INT;
	i2 :	INT;
	i3 :	INT;
	state :	INT;
	domain_copy :	STRING;
	activate_last :	BOOL;
	url_length :	INT;
	char :	BYTE;
	char_count :	INT;
	tid :	BYTE;
	anc :	INT;
	x :	BYTE;
	rr_stop :	BOOL;
	ttl_last :	DWORD;
	ttl_tmp :	DWORD;
	z :	INT;
END_VAR

(*Group:Default*)

VAR_IN_OUT
	IP_C :	oscat_IP_C;(*IP_Control Verwaltungsstruktur*)
	S_BUF :	oscat_NETWORK_BUFFER;
	R_BUF :	oscat_NETWORK_BUFFER;
END_VAR

VAR_INPUT
	ACTIVATE :	BOOL;
	DOMAIN :	STRING;
	IP4_DNS :	DWORD;
END_VAR

VAR_OUTPUT
	IP4 :	DWORD;
	DONE :	BOOL;
	ERROR :	DWORD;
END_VAR

(*@KEY@: WORKSHEET
NAME: DNS_CLIENT
IEC_LANGUAGE: ST
*)
(* Domain Name System (query) *)

CASE state OF

00:	IF ACTIVATE AND NOT activate_last THEN (* auf positive Flanke GET warten *)
		DONE := FALSE;
		ERROR := DWORD#0;
		state := 5;
	END_IF;

05: (* prüfe ob domain schon eine IP4-Adresse ist *)
    IP4_DECODE(str:=DOMAIN);
    IP4 := IP4_DECODE.IP4_DECODE; (* IP4 Adresse direkt weitergeben *)
	IF IP4 > DWORD#00 THEN
		DONE := TRUE;
		state := 0;
        (*####################  DEBUG-MESSAGE  ###################################*)
        (*IF _debug_enable THEN
            LOG_CL.NEW_MSG := 'DNS: S05 IP4 ~1';
            LOG_CL.PRINTF[1]  := DOMAIN;
            LOG_MSG();
        END_IF;*)
        (*########################################################################*)
	ELSE
		ip_state := BYTE#1;
		ttl_last := DWORD#0;
		domain_copy := DOMAIN; (* DOMAIN String sichern *)
		state := 10;
        (*####################  DEBUG-MESSAGE  ###################################*)
        (*IF _debug_enable THEN
            LOG_CL.NEW_MSG := 'DNS: S05 START';
            LOG_MSG();
        END_IF;*)
        (*########################################################################*)
	END_IF;

10:	IF ip_state = BYTE#3 THEN (* Bei IP_Control anmelden *)
		url_length := LEN(domain_copy);
		char_count := 17 + url_length; (* sendebuffer initialisieren *)
		FOR i := 0 TO char_count DO
			S_BUF.BUFFER[i] := BYTE#00;
		END_FOR;
		tid := UINT_TO_BYTE(BYTE_TO_UINT(tid) + UINT#1);
		S_BUF.BUFFER[01] := tid; (* Transaction ID lowbyte *)
		S_BUF.BUFFER[02] := BYTE#16#01; (* Flags: highbyte *)
		S_BUF.BUFFER[05] := BYTE#16#01; (* Questions: lowbyte *)
		i := url_length + 12; (* den servernamen von hinten nach vorne bearbeiten *)
		char_count := 0;
		WHILE i > 12 DO
			CODE(STR:=domain_copy,POS:=i - 12);
			char := CODE.CODE;
			IF char = BYTE#46 THEN (* prüfe auf haupt/sub domänen namens-teiler "." *)
				S_BUF.BUFFER[i] := INT_TO_BYTE(char_count); (* anstelle des teilers "." wird die länge des erkannten haupt/sub domänennames eingetragen *)
				char_count := 0;
			ELSE
				S_BUF.BUFFER[i] := char; (* char in buffer eintragen *)
				char_count := char_count + 1; (* anzahl char zählen *)
			END_IF;
			i := i - 1;
		END_WHILE;
		S_BUF.BUFFER[i] := INT_TO_BYTE(char_count); (* längenangabe des ganz linken (ersten) domänennamens eintragen *)
		i := url_length + 15; (* position hinter dem servernamen *)
		S_BUF.BUFFER[i] := BYTE#01; (* Type: A Hostaddress lowbyte *)
		i := i + 2;
		S_BUF.BUFFER[i] := BYTE#01; (* Class: IN lowbyte *)
		i := i + 1;
		(* IP Datenverkehr einrichten *)
		IP_C.C_PORT := WORD#53; (* Portnummer eintragen *)
		IP_C.C_IP := IP4_DNS; (* IP eintragen *)
		IP_C.C_MODE := BYTE#1; (* Mode: UDP+AKTIV+PORT+IP *)
		IP_C.C_ENABLE := TRUE; (* Verbindungsaufbau freigeben *)
		IP_C.TIME_RESET := TRUE; (* Zeitueberwachung rücksetzen *)
		IP_C.R_OBSERVE  := TRUE; (* Datenempfang ueberwachen *)
		S_BUF.SIZE := INT_TO_UINT(i); (* sendelänge eintragen *)
		R_BUF.SIZE := UINT#0; (* Empfangslänge rücksetzen *)
		state := 30;

        (*####################  DEBUG-MESSAGE  ###################################*)
        (*IF _debug_enable THEN
            LOG_CL.NEW_MSG := 'DNS: S10 SEND';
            LOG_MSG();
        END_IF;*)
        (*########################################################################*)
	END_IF;

30:	IF IP_C.ERROR <> DWORD#00 THEN
		ERROR := IP_C.ERROR;
		state := 99;
        (*####################  DEBUG-MESSAGE  ###################################*)
        (*IF _debug_enable THEN
            LOG_CL.NEW_MSG := 'DNS: S30 ERROR ~1';
            LOG_CL.PRINTF[1]  := DWORD_TO_STRING(ERROR,'%08X');
            LOG_MSG();
        END_IF;*)
        (*########################################################################*)

	ELSIF (S_BUF.SIZE = UINT#0) AND (tid = R_BUF.BUFFER[1]) AND (R_BUF.SIZE >= INT_TO_UINT(34 + url_length)) THEN	(* prüfe ob antwort telegramm die richtige Transaction-ID und mindestlänge hat *)
		ERROR := BYTE_TO_DWORD(R_BUF.BUFFER[3] AND BYTE#2#0000_1111); (* prüfe Return code der Flags. 4 bits *)
		IF ERROR = DWORD#00 THEN
			anc := _BYTE_TO_INT(R_BUF.BUFFER[7]); (* Anzahl der Answer-RR *)
			IP_C.R_OBSERVE := FALSE; (* Datenempfang ueberwachen *)
			state := 40;
		ELSE
			state := 99;
		END_IF;
	END_IF;

40:	IF anc > 0 THEN
		anc := anc - 1;
		z := UINT_TO_INT(R_BUF.SIZE);
		WHILE i < z DO
			x := R_BUF.BUFFER[i];
			IF rr_stop = FALSE THEN
				IF x > BYTE#63 THEN (* zeiger auf namen *)
					i := i + 1;
					rr_stop := TRUE;
				ELSIF x= BYTE#0 THEN (* namens ende *)
					rr_stop := TRUE;
				ELSE
					i := i + _BYTE_TO_INT(x); (* namen *)
				END_IF;
				i := i + 1;
			ELSE
				rr_stop := FALSE;
				i1 := i + 1;
				i3 := i + 3;
				IF R_BUF.BUFFER[i1] = BYTE#1 AND R_BUF.BUFFER[i3] = BYTE#1 THEN (* Type A / Class IN *)
					i := i + 4;
					i1 := i + 1;
					i2 := i + 2;
					i3 := i + 3;
					ttl_tmp := DWORD_OF_BYTE(R_BUF.BUFFER[i],R_BUF.BUFFER[i1],R_BUF.BUFFER[i2],R_BUF.BUFFER[i3]); (* Time to live *)
					i := i + 6;
					IF ttl_tmp >= ttl_last THEN (* TTL ist länger *)
						ttl_last := ttl_tmp;
						i1 := i + 1;
						i2 := i + 2;
						i3 := i + 3;
						IP4 := DWORD_OF_BYTE(R_BUF.BUFFER[i],R_BUF.BUFFER[i1],R_BUF.BUFFER[i2],R_BUF.BUFFER[i3]); (* IP-Adresse *)
					END_IF;
					i := i + 4;
				ELSE
					i := i + 9;
					i := i + _BYTE_TO_INT(R_BUF.BUFFER[i]) + 1; (* offset zu nächsten Block *)
				END_IF;
				EXIT;
			END_IF;
		END_WHILE;
	ELSE
		IF IP4 > DWORD#0 THEN (* gültige RR mit IP gefunden *)
			DONE := TRUE;
            (*####################  DEBUG-MESSAGE  ###################################*)
            (*IF _debug_enable THEN
                LOG_CL.NEW_MSG       := 'DNS: S40 OK';
                LOG_MSG();
            END_IF;*)
            (*########################################################################*)
		ELSE
			ERROR := DWORD#255; (* Daten fehlerhaft - keine IP-Adresse gefunden *)
		END_IF;
		state := 99;
	END_IF;

99:	R_BUF.SIZE := UINT#0; (* Empfangslänge rücksetzen *)
	ip_state := BYTE#4; (* Abmelden *)
	state := 00;

END_CASE;

activate_last := ACTIVATE; (* letzten Status sichern zur Flankenerkennung *)

IP_FIFO(FIFO:=IP_C.FIFO,STATE:=ip_state,ID:=ip_id); (* IP_FIFO *)
IP_C.FIFO:=IP_FIFO.FIFO;
ip_state := IP_FIFO.STATE;
ip_id:=IP_FIFO.ID;

(* revision history

ks	18. oct. 2008	rev 1.0
	original version

ks	20. oct. 2009	rev 1.1
	unbenutzten code entfernt, all buffer base 0

ks	20. dec. 2010	rev 1.2
	parsing nach rfc1305

ks	26. jul. 2011	rev 1.3
	verbesserte ip-auswertung, neue fehlermeldung
*)

(*----------------------------------------------------------------------------------------------------------------*)
(* Flags: 0x0100 (Standard query)                                                                                            *)
(* 0... .... .... .... = Response: Message is a query                                                                   *)
(* .000 0... ....  = Opcode: Standard query (0)                                                                          *)
(* .... ..0. .... .... = Truncated: Message is not truncated                                                          *)
(* .... ...1 .... .... = Recursion desired: Do query recursively                                                    *)
(* .... .... .0.. .... = Z: reserved (0)                                                                                                  *)
(* .... .... ...0 .... = Non-authenticated data OK: Non-authenticated data is unacceptable *)
(*-----------------------------------------------------------------------------------------------------------------*)

(*      0  1  2  3  4  5  6  7  8  9  0  1  2  3  4  5  *)
(*    +--+--+--+--+--+--+--+--+--+--+--+--+--+--+--+--+ *)
(*    |                      ID                       | idx: 0/1   *)
(*    +--+--+--+--+--+--+--+--+--+--+--+--+--+--+--+--+ *)
(*    |QR|   Opcode  |AA|TC|RD|RA|   Z    |   RCODE   | idx: 2/3   *)
(*    +--+--+--+--+--+--+--+--+--+--+--+--+--+--+--+--+ *)
(*    |                    QDCOUNT                    | idx: 4/5   *)
(*    +--+--+--+--+--+--+--+--+--+--+--+--+--+--+--+--+ *)
(*    |                    ANCOUNT                    | idx: 6/7   *)
(*    +--+--+--+--+--+--+--+--+--+--+--+--+--+--+--+--+ *)
(*    |                    NSCOUNT                    | idx: 8/9   *)
(*    +--+--+--+--+--+--+--+--+--+--+--+--+--+--+--+--+ *)
(*    |                    ARCOUNT                    | idx: 10/11 *)
(*    +--+--+--+--+--+--+--+--+--+--+--+--+--+--+--+--+ *)

(*
Errorcodes  Description	References
000	No error. 		 	The request completed successfully.
001	Format error. 		The name server was unable to interpret the query.
002	Server failure.  	The name server was unable to process this query due to a problem with the name server.
003	Name Error. 	 	Meaningful only for responses from an authoritative name server, this code signifies that the domain name referenced in the query does not exist.
004	Not Implemented. 	The name server does not support the requested kind of query.
005	Refused. 			The name server refuses to perform the specified operation for policy reasons.
  						 For example, a name server may not wish to provide the information to the particular requester, or a name server may not wish to perform a particular operation (e.g., zone transfer) for particular data.
006	YXDomain.			Name Exists when it should not.
007	YXRRSet. RR			Set Exists when it should not.
008	NXRRSet. RR			Set that should exist does not.
009	NotAuth.			Server Not Authoritative for zone.
010	NotZone,			Name not contained in zone.
255	Timeout				No Response

beispiel einer DNS Request von google.at
ein request mit 3 Answer-Blocks

Domain Name System (response)
[Request In: 3]
[Time: 0.027533000 seconds]
Transaction ID: 0x5e1a
Flags: 0x8180 (Standard query response, No error)
1... .... .... .... = Response: Message is a response
.000 0... .... .... = Opcode: Standard query (0)
.... .0.. .... .... = Authoritative: Server is not an authority for domain
.... ..0. .... .... = Truncated: Message is not truncated
.... ...1 .... .... = Recursion desired: Do query recursively
.... .... 1... .... = Recursion available: Server can do recursive queries
.... .... .0.. .... = Z: reserved (0)
.... .... ..0. .... = Answer authenticated: Answer/authority portion was not authenticated
.... .... .... 0000 = Reply code: No error (0)
Questions: 1
Answer RRs: 3
Authority RRs: 0
Additional RRs: 0

Queries
google.at: type A, class IN
Name: google.at
Type: A (Host address)
Class: IN (0x0001)

Answers
google.at: type A, class IN, addr 72.14.221.104
Name: google.at
Type: A (Host address)
Class: IN (0x0001)
Time to live: 19 minutes, 9 seconds
Data length: 4
Addr: 72.14.221.104

google.at: type A, class IN, addr 66.249.93.104
Name: google.at
Type: A (Host address)
Class: IN (0x0001)
Time to live: 19 minutes, 9 seconds
Data length: 4
Addr: 66.249.93.104

google.at: type A, class IN, addr 216.239.59.104
Name: google.at
Type: A (Host address)
Class: IN (0x0001)
Time to live: 19 minutes, 9 seconds
Data length: 4
Addr: 216.239.59.104
*)

(*@KEY@: END_WORKSHEET *)
END_FUNCTION_BLOCK

(* ---- DNS_REV_CLIENT.ST ---- *)
(*@PROPERTIES_EX@
TYPE: POU
LOCALE: 0
IEC_LANGUAGE: ST
PLC_TYPE: independent
PROC_TYPE: independent
GROUP: NETWORK
*)
(*@KEY@:DESCRIPTION*)
version 1.0	28. dec. 2009
programmer 	ks
tested BY	ks

DNS_REV_CLIENT führt eine Reverse-Domain-Name Abfrage durch, und ermittelt aus einer IP-Adresse den zugehörigen Domain-Namen.

(*@KEY@:END_DESCRIPTION*)
FUNCTION_BLOCK DNS_REV_CLIENT

(*Group:Default*)

VAR_IN_OUT
	IP_C :	oscat_IP_C;(*IP_Control Verwaltungsstruktur*)
	S_BUF :	oscat_NETWORK_BUFFER;
	R_BUF :	oscat_NETWORK_BUFFER;
END_VAR

VAR_INPUT
	ACTIVATE :	BOOL;
	IP4 :	DWORD;
	IP4_DNS :	DWORD;
END_VAR

VAR_OUTPUT
	DOMAIN :	STRING;
	DONE :	BOOL;
	ERROR :	DWORD;
END_VAR

VAR
	IP_FIFO :	IP_FIFO;
	ip_state :	BYTE;
	ip_id :	BYTE;
	state :	INT;
	ip4_copy :	DWORD;
	d :	oscat_STRING27;
	activate_last :	BOOL;
	i :	INT;
	dl :	INT;
	p1 :	INT;
	char :	BYTE;
	char_count :	INT;
	tid :	BYTE;
	BUFFER_TO_STRING :	BUFFER_TO_STRING_NW;
	CODE :	CODE;
END_VAR

(*@KEY@: WORKSHEET
NAME: DNS_REV_CLIENT
IEC_LANGUAGE: ST
*)
(* Domain Name System (query) *)

CASE state OF
00: (* auf positive Flanke GET warten *)
	IF ACTIVATE AND NOT activate_last THEN
		ERROR := DWORD#0;
		ip4_copy := ip4; (* IP4 sichern *)
		ip_state := BYTE#1;
		DOMAIN := '';
		DONE := FALSE;

		d := '';
		FOR i := 1 TO 4 DO
			d := CONCAT(d,BYTE_TO_STRING(DWORD_TO_BYTE(IP4),'%u'));
			d := CONCAT(d,'.');
			IP4 := ROR(IP4,8);
		END_FOR;
		d := CONCAT(d,'in-addr.arpa');
		state := 10;
	END_IF;

10: (* Bei IP_Control anmelden *)
	IF ip_state = BYTE#3 THEN
		dl := LEN(d);

		(* sendebuffer initialisieren *)
		char_count := 17 + dl;
		FOR i := 0 TO char_count DO
			S_BUF.BUFFER[i] := BYTE#00;
		END_FOR;

		tid := UINT_TO_BYTE(BYTE_TO_UINT(tid) + UINT#1);
		S_BUF.BUFFER[01] := tid; (* Transaction ID lowbyte *)
		S_BUF.BUFFER[02] := BYTE#16#01; (* Flags: highbyte *)
		S_BUF.BUFFER[05] := BYTE#16#01; (* Questions: lowbyte *)

		(* den servernamen von hinten nach vorne bearbeiten *)
		i := dl + 12;
		char_count := 0;

		WHILE i > 12 DO
			CODE(STR:=d,POS:=i - 12);
			char:=CODE.CODE;

			(* prüfe auf haupt/sub domänen namens-teiler "." *)
			IF char = BYTE#46 THEN
				(* anstelle des teilers "." wird die länge des erkannten haupt/sub domänennames eingetragen *)
				S_BUF.BUFFER[i] := INT_TO_BYTE(char_count);
				char_count := 0;
			ELSE
				S_BUF.BUFFER[i] := char; (* char in buffer eintragen *)
				char_count := char_count + 1; (* anzahl char zählen *)
			END_IF;
			i := i - 1;
		END_WHILE;

		S_BUF.BUFFER[i] := INT_TO_BYTE(char_count); (* längenangabe des ganz linken (ersten) domänennamens eintragen *)
		i := dl + 15; (* position hinter dem servernamen *)
		S_BUF.BUFFER[i] := BYTE#12; (* Type: PTR (Domain name pointer) lowbyte *)
		i := i + 2;
		S_BUF.BUFFER[i] := BYTE#01; (* Class: IN lowbyte *)
		i := i + 1;

		(* IP Datenverkehr einrichten *)
		IP_C.C_PORT := WORD#53; (* Portnummer eintragen *)
		IP_C.C_IP := IP4_DNS; (* IP eintragen *)
		IP_C.C_MODE := BYTE#1; (* Mode: UDP+AKTIV+PORT+IP *)
		IP_C.C_ENABLE := TRUE; (* Verbindungsaufbau freigeben *)
		IP_C.TIME_RESET := TRUE; (* Zeitueberwachung rücksetzen *)
		IP_C.R_OBSERVE  := TRUE; (* Datenempfang ueberwachen *)
		S_BUF.SIZE := INT_TO_UINT(i); (* sendelänge eintragen *)
		R_BUF.SIZE := UINT#0; (* Empfangslänge rücksetzen *)
		state := 30;
	END_IF;

30:
	IF IP_C.ERROR <> DWORD#00 THEN
		ERROR := IP_C.ERROR;
	(* prüfe ob antwort telegramm die richtige Transaction-ID und mindestlänge hat *)
	ELSIF (S_BUF.SIZE = UINT#0) AND (tid = R_BUF.BUFFER[1]) AND (R_BUF.SIZE >= INT_TO_UINT(i+12)) THEN

		(* prüfe Return code der Flags. 4 bits *)
		ERROR := BYTE_TO_DWORD(R_BUF.BUFFER[3] AND BYTE#2#0000_1111);

		IF ERROR = DWORD#00 THEN

			i := UINT_TO_INT(R_BUF.SIZE) - 2;
			WHILE R_BUF.BUFFER[i] > BYTE#0 DO
				IF i = 0 THEN EXIT; END_IF;
				i := i - 1;
			END_WHILE;

			i := i + 2;
			p1 := i + 1;
			WHILE i < UINT_TO_INT(R_BUF.SIZE) DO
				dl := _BYTE_TO_INT(R_BUF.BUFFER[i]);
				IF dl > 0 THEN
					R_BUF.BUFFER[i] := BYTE#46;
					i := i + dl + 1;
				ELSE

					BUFFER_TO_STRING(PT:=R_BUF.BUFFER,SIZE:=UINT#4096,START:=INT_TO_UINT(p1),STOP:=INT_TO_UINT(i-1));
					R_BUF.BUFFER:=BUFFER_TO_STRING.PT;
					DOMAIN:=BUFFER_TO_STRING.BUFFER_TO_STRING;
					EXIT;
				END_IF;
			END_WHILE;
			state := 0;
			DONE := TRUE;
		END_IF;
	END_IF;

	IF ERROR <> DWORD#0 THEN
		state := 0;
	END_IF;

	IF state = 0 THEN
		IP_C.R_OBSERVE := FALSE; (* Datenempfang ueberwachen *)
		ip_state := BYTE#4; (* Abmelden *)
	END_IF;

END_CASE;

activate_last := ACTIVATE; (* letzten Status sichern zur Flankenerkennung *)

(* IP_FIFO *)
IP_FIFO(FIFO:=IP_C.FIFO,STATE:=ip_state,ID:=ip_id);
IP_C.FIFO:=IP_FIFO.FIFO;
ip_state:=IP_FIFO.STATE;
ip_id:=IP_FIFO.ID;

(* revision history

ks	28. dec. 2009	rev 1.0
	original version

*)

(*----------------------------------------------------------------------------------------------------------------*)
(* Flags: 0x0100 (Standard query)                                                                                            *)
(* 0... .... .... .... = Response: Message is a query                                                                   *)
(* .000 0... ....  = Opcode: Standard query (0)                                                                          *)
(* .... ..0. .... .... = Truncated: Message is not truncated                                                          *)
(* .... ...1 .... .... = Recursion desired: Do query recursively                                                    *)
(* .... .... .0.. .... = Z: reserved (0)                                                                                                  *)
(* .... .... ...0 .... = Non-authenticated data OK: Non-authenticated data is unacceptable *)
(*-----------------------------------------------------------------------------------------------------------------*)

(*
Errorcodes  Description	References
000	No error. 		 	The request completed successfully.
001	Format error. 		The name server was unable to interpret the query.
002	Server failure.  	The name server was unable to process this query due to a problem with the name server.
003	Name Error. 	 	Meaningful only for responses from an authoritative name server, this code signifies that the domain name referenced in the query does not exist.
004	Not Implemented. 	The name server does not support the requested kind of query.
005	Refused. 			The name server refuses to perform the specified operation for policy reasons.
  						 For example, a name server may not wish to provide the information to the particular requester, or a name server may not wish to perform a particular operation (e.g., zone transfer) for particular data.
006	YXDomain.			Name Exists when it should not.
007	YXRRSet. RR			Set Exists when it should not.
008	NXRRSet. RR			Set that should exist does not.
009	NotAuth.			Server Not Authoritative for zone.
010	NotZone,			Name not contained in zone.
255	Timeout				No Response
*)

(*@KEY@: END_WORKSHEET *)
END_FUNCTION_BLOCK

(* ---- FILE_BLOCK.ST ---- *)
(*@PROPERTIES_EX@
TYPE: POU
LOCALE: 0
IEC_LANGUAGE: ST
PLC_TYPE: independent
PROC_TYPE: independent
GROUP: FILE
*)
(*@KEY@:DESCRIPTION*)
version 1.0		23. sep. 2010
programmer 		ks
tested by		ks

FILE_BLOCK liefert das angeforderte Byte einer Datei durch einlesen von möglichst grossen Datenblöcken

(*@KEY@:END_DESCRIPTION*)
FUNCTION_BLOCK FILE_BLOCK

(*Group:parameter*)

VAR_IN_OUT
	MODE :	BYTE;
	FILENAME :	STRING;
	FSD :	oscat_FILE_SERVER_DATA;
	PT :	oscat_NETWORK_BUFFER;
END_VAR

VAR_INPUT
	POS :	UDINT;
END_VAR

VAR_OUTPUT
	ERROR :	BYTE;
	DATA :	BYTE;
END_VAR

(*Group:log*)

VAR
	(*<LOG_MSG :	LOG_MSG;>*)
	(*<_debug_enable :	BOOL := TRUE;>*)
END_VAR

VAR_EXTERNAL
	(*<LOG_CL :	us_LOG_CONTROL;>*)
END_VAR

(*Group:var*)

VAR
	step :	INT;
	i :	INT;
	data_start :	UDINT;
	data_stop :	UDINT;
END_VAR

(*@KEY@: WORKSHEET
NAME: FILE_BLOCK
IEC_LANGUAGE: ST
*)
CASE step OF
0:	IF MODE > BYTE#0 THEN
		ERROR := BYTE#0;
		IF FSD.FILE_OPEN AND (FSD.FILE_SIZE = UDINT#0 OR POS >= FSD.FILE_SIZE) THEN
			ERROR := BYTE#255;
			MODE := BYTE#0;
		ELSIF POS < data_start OR POS > data_stop OR NOT FSD.FILE_OPEN THEN (* Daten lesen notwendig *)
			FSD.FILENAME := FILENAME;
			FSD.MODE := BYTE#1; (* open + read *)
			FSD.OFFSET := POS;
			PT.SIZE := UINT#65535; (* maximale anzahl lesen *);
			data_start := UDINT#0;
			data_stop := UDINT#0;
			step := 10;
		ELSE (* Daten sind im Buffer vorhanden *)
			i := UDINT_TO_INT(POS - data_start); (* index berechnen *)
			DATA := PT.BUFFER[i];
			MODE := BYTE#0;
			(* ---------------------- Debug-Message ----------------------------*)
			(*IF _debug_enable THEN
				LOG_CL.NEW_MSG := 'FB: Pos: ~1 Byte: ~2 >~3<';
				LOG_CL.PRINTF[1] := UDINT_TO_STRING(POS,'%03u');
				LOG_CL.PRINTF[2] := BYTE_TO_STRING(DATA,'%03u');
				LOG_CL.PRINTF[3] := BYTE_TO_STRING(DATA,'%c');
				LOG_MSG();
			END_IF;*)
			(* -----------------------------------------------------------------*)
		END_IF;
	END_IF;

10:	IF FSD.MODE = BYTE#0 THEN (* Befehl beendet *)
		IF FSD.ERROR > BYTE#0 THEN
			ERROR := FSD.ERROR; (* Fehler ausgeben *)
			MODE := BYTE#0;
		ELSE
			data_start := POS;
			data_stop := POS + UINT_TO_UDINT(PT.SIZE) - UDINT#1;
		END_IF;
		step := 0;
	END_IF;
END_CASE;

(* revision history
ks	23. sep. 2010	rev 1.0
	original version
*)

(*@KEY@: END_WORKSHEET *)
END_FUNCTION_BLOCK

(* ---- FILE_SERVER.ST ---- *)
(*@PROPERTIES_EX@
TYPE: POU
LOCALE: 0
IEC_LANGUAGE: ST
PLC_TYPE: independent
PROC_TYPE: independent
GROUP: HARDWARE
*)
(*@KEY@:DESCRIPTION*)
version 1.0		23. sep. 2010
programmer 		ks
tested by		ks

FILE_SERVER ermöglicht den Zugriff auf Dateien mittels Plattform-Neutraler Schnittstelle

Befehle:
1 = File_Open_Exist + File_Read
2 = File_Open_Exist + File_Write
3 = File_Open_New   + File_Write
4 = File_Remove
5 = File_Close

- Action -
1 = file_open   (open)
2 = file_close  (close)
3 = file_read   (read)
4 = file_write  (write)
5 = file_seek   (setpos)
6 = file_tell   (getpos)
7 = file_remove (delete)

---- fehlermeldungen----

000 (00) kein Fehler

002 (02) file_open - Die maximale Anzahl von Dateien ist bereits geöffnet.
004 (04) file_open - Die Datei ist bereits geöffnet.
005 (05) file_open - Die Datei ist schreibgeschützt oder Zugriff verweigert.
006 (06) file_open - Dateiname nicht angegeben.

011 (01) file_close - Ungültiger Dateihandle.
030 (20) file_close - Datei konnte nicht geschlossen werden.

041 (01) file_read - Ungültiger Dateihandle.
050 (10) file_read - Dateiende erreicht.
052 (12) file_read - Die Anzahl der zu lesenden Zeichen ist größer als der Datenpuffer.
062 (22) file_read - Es konnten keine Daten gelesen werden.

071 (01) file_write - Ungültiger Dateihandle.
081 (11) file_write - Es ist kein Speicher zum Schreiben der Daten verfügbar.
082 (12) file_write - Die Anzahl der zu schreibenden Zeichen ist größer als der Datenpuffer.
093 (23) file_write - Es konnten keine Daten geschrieben werden.

101 (01) file_seek - Ungültiger Dateihandle.
113 (13) file_seek - Ungültiger Positionierungsmodus oder die angegebene Position liegt vor dem Dateianfang.
124 (24) file_seek - Die Position konnte nicht gesetzt werden.

131 (01) file_tell - Ungültiger Dateihandle.

142 (02) file_remove - Die maximale Anzahl von Dateien ist bereits geöffnet.
143 (03) file_remove - Die Datei konnte nicht gefunden werden.
145 (05) file_remove - Die Datei ist geöffnet, schreibgeschützt oder Zugriff verweigert.
146 (06) file_remove - Dateiname nicht angegeben.
161 (21) file_remove - Datei konnte nicht gelöscht werden.

255: Position liegt hinter dem Dateiende (Applikationserror)

(*@KEY@:END_DESCRIPTION*)
FUNCTION_BLOCK FILE_SERVER

(*Group:neu*)

VAR
	buf_size :	UDINT := UDINT#4096;
	handle :	UINT;(*Filehandle*)
	read_max_length :	UDINT;(*maximale Datenlänge*)
	file_position :	UDINT;(*aktueller Schreib/Lesezeiger*)
	used_filename :	STRING;(*aktueller Dateiname*)
	close_time :	TIME;
	length_read :	UDINT;
	write_length :	UDINT;
	length_written :	UDINT;
	open_handle :	UINT;
	seek_mode :	UINT;
	seek_position :	UDINT;
	tell_position :	UDINT;
END_VAR

(*Group:lokal*)

VAR
	last_mode :	BYTE;
	command :	BYTE;
	error_code :	BYTE;
	error :	BOOL;
	file_change :	BOOL;
	step :	INT;
	t_diff :	TIME;
	tx_last :	TIME;
	tx :	TIME;
END_VAR

(*Group:parameter*)

VAR_IN_OUT
	FSD :	oscat_FILE_SERVER_DATA;
	PT :	oscat_NETWORK_BUFFER;
END_VAR

(*Group:log*)

VAR
	(*<_debug_enable :	BOOL := TRUE;>*)
	(*<step_last :	INT;>*)
	(*<LOG_MSG :	LOG_MSG;>*)
END_VAR

VAR_EXTERNAL
	(*<LOG_CL :	us_LOG_CONTROL;>*)
END_VAR

(*Group:Instance*)

VAR
	FILE_REMOVE :	FILE_REMOVE;
	FILE_OPEN :	FILE_OPEN;
	FILE_SEEK :	FILE_SEEK;
	FILE_TELL :	FILE_TELL;
	FILE_CLOSE :	FILE_CLOSE;
	FILE_READ :	FILE_READ;
	FILE_WRITE :	FILE_WRITE;
	T_PLC_MS :	T_PLC_MS;
END_VAR

(*@KEY@: WORKSHEET
NAME: FILE_SERVER
IEC_LANGUAGE: ST
*)
(* read system timer *)
T_PLC_MS();
tx := UDINT_TO_TIME(T_PLC_MS.T_PLC_MS);
t_diff := tx - tx_last;
tx_last := tx;

CASE step OF
0:
	IF FSD.MODE = LIMIT(BYTE#1,FSD.MODE,BYTE#5) THEN
   		(* ---------------------- Debug-Message ----------------------------*)
		(*IF _debug_enable THEN
			LOG_CL.NEW_MSG := 'File_Start Mode=~1';
			LOG_CL.PRINTF[1] := BYTE_TO_STRING (FSD.MODE,'%u');
			LOG_MSG();
		END_IF;*)
		(* -----------------------------------------------------------------*)
		close_time := T#1ms; (* wenn Schritt aktiv ist, dann Close-Timer rücksetzen *)
		IF handle = UINT#00 AND FSD.MODE <= BYTE#3 THEN (* Mode 1,2,3 und file nicht geöffnet *)
			step := 100; (* File muss erst geöffnet werden *)
		ELSE
			(* File ist schon geöffnet - alten und neuen Filenamen vergleichen *)
			IF EQ_STRING(used_filename, FSD.FILENAME) AND FSD.MODE = last_mode THEN (* kein Moduswechsel ? *)
				step := 200; (* ohne open prozedure weitermachen *)
			ELSE
				step := 32000; (* (* mode 3,4,5 - File_Close ausführen *)
				file_change := FSD.MODE <> BYTE#5; (* mode 5 - File_close ausschliessen *)
			END_IF;
		END_IF;
	ELSIF handle > UINT#0 THEN (* offene Datei gefunden - AutoClose Modus *)
		IF FSD.AUTO_CLOSE > T#0s THEN
			close_time := close_time + t_diff; (* Close_Time hochzählen *)
			IF close_time > FSD.AUTO_CLOSE THEN (* Zeit überschrittenen *)
				step := 32000; (* automatisch Datei schliessen *)
			END_IF;
		END_IF;
	END_IF;

100:
	IF FSD.MODE = BYTE#3 OR FSD.MODE = BYTE#4 THEN
		command := BYTE#7; (* File Remove *)
		step := 110;
	ELSE
		step := 120; (* File Open ausführen *)
	END_IF;

110: (* File Remove *)
	IF command = BYTE#0  THEN
		IF (FSD.MODE = BYTE#4) OR (error and error_code <> BYTE#143) THEN (* Mode: File Remove *)
			step := 30000; (* Beenden *)
		ELSE
			step := 120;
		END_IF;
	END_IF;

120:
	command := BYTE#1; (* File Open *)
	last_mode := FSD.MODE;
	step := 122;

122: (* File Open *)
	IF command = BYTE#0 THEN
		IF error THEN
			step := 30000; (* Beenden *)
		ELSE
			(* Filedaten eintragen *)
			close_time := T#1ms; (* Timer freigeben *)
			handle := open_handle;
			used_filename := FSD.FILENAME;
			file_position := UDINT#4294967295; (* maximal = unbekannt *)
			FSD.FILE_SIZE := UDINT#0;
			step := 125;
		END_IF;
	END_IF;

125: (* File Seek - Dateigroesse bestimmen *)
	seek_mode := UINT#2;  (* Positionierung relativ zum Dateiende *)
	seek_position := UDINT#0;
	command := BYTE#5; (* File Seek *)
	step := 130;

130: (* File Seek *)
	IF command = BYTE#0 THEN
		IF Error THEN
			step := 30000; (* Beenden *)
		ELSE
			step := 140;
		END_IF;
	END_IF;

140: (* File Tell - Position des Schreib/Lesezeiger auslesen *)
	command := BYTE#6; (* File Tell *)
	step := 150;

150: (* File Tell *)
	IF command = BYTE#0 THEN
		IF Error THEN
			step := 30000; (* Beenden *)
		ELSE
			FSD.FILE_SIZE := tell_position; (* aktuelle Dateigroesse *)
			file_position := tell_position;
			FSD.FILE_OPEN := TRUE;
			step := 200;
		END_IF;
	END_IF;

200: (* File Seek *)
	IF FSD.OFFSET > FSD.FILE_SIZE THEN (* prüfe auf gültige offset-vorgabe *)
		error_code := BYTE#255;
		step := 30000; (* Beenden *)
	ELSIF FSD.OFFSET <> file_position THEN
		command := BYTE#5; (* File-Seek *)
		seek_mode := UINT#0; (* Positionierung relativ zum Dateianfang *)
		seek_position := FSD.OFFSET;
		step := 210;
	ELSE
		step := 300;
	END_IF;

210: (* File Seek *)
	IF command = BYTE#0 THEN
		file_position := seek_position;
		IF Error THEN
			step := 30000; (* Beenden *)
		ELSE
			step := 300;
		END_IF;
	END_IF;

300:
	IF FSD.MODE = BYTE#1 THEN
		step := 400; (* Read *)
	ELSE
		step := 500; (* Write *)
	END_IF;

400: (* File Read *)
	IF UINT_TO_UDINT(PT.SIZE) > buf_size THEN (* Leselänge auf Buffergroesse begrenzen *)
		read_max_length := buf_size;
	ELSE
		read_max_length := UINT_TO_UDINT(PT.SIZE);
	END_IF;

	(* Leselänge an Dateilänge anpassen *)
	IF file_position + read_max_length > FSD.FILE_SIZE THEN
		read_max_length := FSD.FILE_SIZE - file_position;
	END_IF;

	IF read_max_length > UDINT#0 THEN
		command := BYTE#3; (* File_Read *)
		step := INT#410;
	ELSE
		PT.SIZE := UINT#0;
		step := 30000; (* Beenden *)
	END_IF;

410: (* File Read *)
	IF command = BYTE#0 THEN
		PT.SIZE := UDINT_TO_UINT(length_read);
		IF NOT Error THEN
			file_position := file_position + length_read; (* aktueller File_Position korrigieren *)
			FSD.OFFSET := file_position;
		END_IF;
		step := 30000; (* Beenden *)
	END_IF;

500: (* File Write *)
	IF UINT_TO_UDINT(PT.SIZE) > buf_size THEN (* Schreiblänge auf Buffergroesse begrenzen *)
		write_length := buf_size;
	ELSE
		write_length := UINT_TO_UDINT(PT.SIZE);
	END_IF;

	IF write_length > UDINT#0 THEN
		command := BYTE#4; (* File_Write *)
		step := INT#510;
	ELSE
		step := 30000; (* Beenden *)
	END_IF;

510:
	IF command = BYTE#0 THEN
		IF NOT Error THEN
			file_position := file_position + length_written; (* aktueller File_Position korrigieren *)
			FSD.OFFSET := file_position;
			IF file_position > FSD.FILE_SIZE THEN (* Datei ist groesser geworden *)
				FSD.FILE_SIZE := file_position;
			END_IF;
		END_IF;
		step := 30000; (* Beenden *)
	END_IF;

(* --------------------------------------------- *)

30000: (* Befehl fertig *)
	FSD.MODE := BYTE#0;
	FSD.ERROR := error_code;
	step := 0;
	(* ---------------------- Debug-Message ----------------------------*)
	(*IF _debug_enable THEN
		LOG_CL.NEW_MSG := 'File_Stop: File ~1, error ~7, code ~8';
		LOG_CL.PRINTF[1]  := used_filename;
		LOG_CL.PRINTF[7]  := INT_TO_STRING(BOOL_TO_INT(error),'%d');
		LOG_CL.PRINTF[8]  := BYTE_TO_STRING(error_code,'%u');
		LOG_MSG();
	END_IF;*)
	(* -----------------------------------------------------------------*)

32000:
	close_time := T#0s; (* Timer stoppen *)
	IF handle > UINT#0 THEN
		command := BYTE#2; (* File_Close ausführen *)
	END_IF;
	step := 32100;

32100:
	IF command = BYTE#0 THEN (* File Close beendet *)
		(* Filedaten ablöschen *)
		FSD.FILE_OPEN := FALSE;
		file_position := UDINT#0;
		FSD.FILE_SIZE := UDINT#0;
		FSD.OFFSET := UDINT#0;
		used_filename := '';
		handle := UINT#00;

		(* File_Name wurde fliegend geändert ? *)
		IF file_change THEN
			file_change := FALSE;
			step := 100;
		ELSE
			step := 30000;
		END_IF;
	END_IF;

END_CASE;

(* ------------ File Open ------------- *)
FILE_OPEN.Execute := command = BYTE#1;
FILE_OPEN.Name := FSD.FILENAME;
FILE_OPEN();
open_handle := FILE_OPEN.Handle;

IF command = BYTE#1 THEN
	IF FILE_OPEN.Done THEN
		error := FILE_OPEN.Error;
		command := BYTE#0;
		error_code := SEL_BYTE(error,BYTE#00,UINT_TO_BYTE(FILE_OPEN.ErrorID));
		(* ---------------------- Debug-Message ----------------------------*)
		(*IF _debug_enable THEN
			LOG_CL.NEW_MSG := 'Open: File ~1, error ~7, code ~8';
			LOG_CL.PRINTF[1] := FSD.FILENAME;
			LOG_CL.PRINTF[7] := INT_TO_STRING(BOOL_TO_INT(error),'%d');
			LOG_CL.PRINTF[8] := BYTE_TO_STRING(error_code,'%u');
			LOG_MSG();
		END_IF;*)
		(* -----------------------------------------------------------------*)
	END_IF;
END_IF;

(* ----------- File Close ------------- *)
FILE_CLOSE.Execute := command = BYTE#2;
FILE_CLOSE.Handle := Handle;
FILE_CLOSE();

IF command = BYTE#2 THEN
	IF FILE_CLOSE.Done THEN
		error := FILE_CLOSE.Error;
		command := BYTE#0;
		error_code := SEL_BYTE(error,BYTE#00,UINT_TO_BYTE(FILE_CLOSE.ErrorID + UINT#10)); (* Errorcode basis verschieben *)
		(* ---------------------- Debug-Message ----------------------------*)
		(*IF _debug_enable THEN
			LOG_CL.NEW_MSG := 'Close: File ~1, error ~7, code ~8';
			LOG_CL.PRINTF[1] := used_filename;
			LOG_CL.PRINTF[7] := INT_TO_STRING(BOOL_TO_INT(error),'%d');
			LOG_CL.PRINTF[8] := BYTE_TO_STRING(error_code,'%u');
			LOG_MSG();
		END_IF;*)
		(* -----------------------------------------------------------------*)
	END_IF;
END_IF;

(* ------------ File Read ------------- *)
FILE_READ.Execute := command = BYTE#3;
FILE_READ.Handle := handle;
FILE_READ.MaxLength := read_max_length;
FILE_READ.Buffer := PT.BUFFER;
FILE_READ();
PT.BUFFER := FILE_READ.Buffer;

IF command = BYTE#3 THEN
	IF FILE_READ.Done THEN
		error := FILE_READ.Error;
		command := BYTE#0;
		length_read :=  FILE_READ.LengthRead;
		error_code := SEL_BYTE(error,BYTE#00,UINT_TO_BYTE(FILE_READ.ErrorID + UINT#40)); (* Errorcode basis verschieben *)
		(* ---------------------- Debug-Message ----------------------------*)
		(*IF _debug_enable THEN
			LOG_CL.NEW_MSG := 'Read: File ~1, soll ~2,ist ~3, offset ~4 ,error ~7, code ~8';
			LOG_CL.PRINTF[1] := used_filename;
			LOG_CL.PRINTF[2] := UDINT_TO_STRING(read_max_length,'%u');
			LOG_CL.PRINTF[3] := UDINT_TO_STRING(length_read,'%u');
			LOG_CL.PRINTF[4] := UDINT_TO_STRING(FSD.OFFSET,'%u');
			LOG_CL.PRINTF[7] := INT_TO_STRING(BOOL_TO_INT(error),'%d');
			LOG_CL.PRINTF[8] := BYTE_TO_STRING(error_code,'%u');
			LOG_MSG();
		END_IF;*)
		(* -----------------------------------------------------------------*)
	END_IF;
END_IF;

(* ------------ File Write ------------- *)
FILE_WRITE.Execute   := command = BYTE#4;
FILE_WRITE.Handle    := handle;
FILE_WRITE.Length    := write_length ;
FILE_WRITE.Buffer    := PT.BUFFER;
FILE_WRITE();
PT.BUFFER := FILE_WRITE.Buffer;

IF command = BYTE#4 THEN
	IF FILE_WRITE.Done THEN
		error := FILE_WRITE.Error;
		command := BYTE#0;
		(*length_written := FILE_WRITE.LengthWritten; Originalcode !! *)
		length_written := write_length; (* Workaround für BUG *)
		error_code := SEL_BYTE(error,BYTE#00,UINT_TO_BYTE(FILE_WRITE.ErrorID + UINT#70)); (* Errorcode basis verschieben *)
		(* ---------------------- Debug-Message ----------------------------*)
		(*IF _debug_enable THEN
			LOG_CL.NEW_MSG := 'Write: File ~1, soll ~2,ist ~3, offset ~4 ,error ~7, code ~8';
			LOG_CL.PRINTF[1] := used_filename;
			LOG_CL.PRINTF[2] := UDINT_TO_STRING(write_length,'%u');
			LOG_CL.PRINTF[3] := UDINT_TO_STRING(length_written,'%u');
			LOG_CL.PRINTF[4] := UDINT_TO_STRING(FSD.OFFSET,'%u');
			LOG_CL.PRINTF[7] := INT_TO_STRING(BOOL_TO_INT(error),'%d');
			LOG_CL.PRINTF[8] := BYTE_TO_STRING(error_code,'%u');
			LOG_MSG();
		END_IF;*)
		(* -----------------------------------------------------------------*)
	END_IF;
END_IF;

(* ------------ File Seek ------------- *)
FILE_SEEK.Execute  := command = BYTE#5;
FILE_SEEK.Handle   := handle;
FILE_SEEK.Mode     := seek_mode;
FILE_SEEK.Position := UDINT_TO_DINT(seek_position);
FILE_SEEK();

IF command = BYTE#5 THEN
	IF FILE_SEEK.Done THEN
		error := FILE_SEEK.Error;
		command := BYTE#0;
		error_code := SEL_BYTE(error,BYTE#00,UINT_TO_BYTE(FILE_SEEK.ErrorID + UINT#100)); (* Errorcode basis verschieben *)
		(* ---------------------- Debug-Message ----------------------------*)
		(*IF _debug_enable THEN
			LOG_CL.NEW_MSG := 'Seek: File ~1, mode ~2,pos ~3 ,error ~7, code ~8';
			LOG_CL.PRINTF[1] := used_filename;
			LOG_CL.PRINTF[2] := UINT_TO_STRING(seek_mode,'%u');
			LOG_CL.PRINTF[3] := UDINT_TO_STRING(seek_position,'%u');
			LOG_CL.PRINTF[7] := INT_TO_STRING(BOOL_TO_INT(error),'%d');
			LOG_CL.PRINTF[8] := BYTE_TO_STRING(error_code,'%u');
			LOG_MSG();
		END_IF;*)
		(* -----------------------------------------------------------------*)
	END_IF;
END_IF;

(* ------------ File Tell ------------- *)
FILE_TELL.Execute := command = BYTE#6;
FILE_TELL.Handle := handle;
FILE_TELL();

IF command = BYTE#6 THEN
	IF FILE_TELL.Done THEN
		error := FILE_TELL.Error;
		command := BYTE#0;
		tell_position := DINT_TO_UDINT(FILE_TELL.Position);
		error_code := SEL_BYTE(error,BYTE#00,UINT_TO_BYTE(FILE_TELL.ErrorID + UINT#130)); (* Errorcode basis verschieben *)
		(* ---------------------- Debug-Message ----------------------------*)
		(*IF _debug_enable THEN
			LOG_CL.NEW_MSG := 'Tell: File ~1, pos ~3 ,error ~7, code ~8';
			LOG_CL.PRINTF[1] := used_filename;
			LOG_CL.PRINTF[3] := UDINT_TO_STRING(tell_position,'%u');
			LOG_CL.PRINTF[7] := INT_TO_STRING(BOOL_TO_INT(error),'%d');
			LOG_CL.PRINTF[8] := BYTE_TO_STRING(error_code,'%u');
			LOG_MSG();
		END_IF;*)
		(* -----------------------------------------------------------------*)
	END_IF;
END_IF;

(* ------------ File Remove ------------- *)
FILE_REMOVE.Execute := command = BYTE#7;
FILE_REMOVE.Name := FSD.FILENAME;
FILE_REMOVE();

IF command = BYTE#7 THEN
	IF FILE_REMOVE.Done THEN
		error := FILE_REMOVE.Error;
		command := BYTE#0;
		error_code := SEL_BYTE(error,BYTE#00,UINT_TO_BYTE(FILE_REMOVE.ErrorID + UINT#140)); (* Errorcode basis verschieben *)
		(* ---------------------- Debug-Message ----------------------------*)
		(*IF _debug_enable THEN
			LOG_CL.NEW_MSG := 'Remove: File ~1, error ~7, code ~8';
			LOG_CL.PRINTF[1] := used_filename;
			LOG_CL.PRINTF[7] := INT_TO_STRING(BOOL_TO_INT(error),'%d');
			LOG_CL.PRINTF[8] := BYTE_TO_STRING(error_code,'%u');
			LOG_MSG();
		END_IF;*)
		(* -----------------------------------------------------------------*)
	END_IF;
END_IF;

(* ---------------------- Debug-Message ----------------------------*)
(*IF _debug_enable THEN
	IF step_last <> step THEN
		LOG_CL.NEW_MSG := 'Step: ~1';
		LOG_CL.PRINTF[1]  := INT_TO_STRING(step,'%d');
		LOG_MSG();
	END_IF;
	step_last := step;
END_IF;*)
(* -----------------------------------------------------------------*)

(* revision history
ks	23. sep. 2010	rev 1.0
	original version
*)

(*@KEY@: END_WORKSHEET *)
END_FUNCTION_BLOCK

(* ---- FTP_CLIENT.ST ---- *)
(*@PROPERTIES_EX@
TYPE: POU
LOCALE: 0
IEC_LANGUAGE: ST
PLC_TYPE: independent
PROC_TYPE: independent
GROUP: NETWORK
*)
(*@KEY@:DESCRIPTION*)
(*
version 1.2		11.may 2011
programmer		ks
tested by		ks

FTP_CLIENT dient zum senden und empfangen von dateien von einem FTP-Server.

110 Restart marker reply 										Markierung für Wiederaufnahme der Übertragung
120 Service ready in x minutes 									Dienst steht in x Minuten zu Verfügung
125 Data connection already open; 								transfer starting Datenverbindung besteht bereits; beginne mit der Übertragung
150 File status okay; about to open data connection 					Dateistatus OK; Datenverbindung wird aufgebaut
200 Command okay 											Befehl OK
202 Command not implemented 									Befehl nicht implementiert
211   														Antwort für Systemstatus oder Hilfefunktion des Systems
212   														Verzeichnisstatus
213   														Dateistatus
214   														Meldung der Hilfefunktion
215 NAME system type 										Angabe des Systemtyps
220 Service ready for new user 									Dienst bereit für neuen Benutzer
221 Service closing control connection 							Steuerverbindung des Dienstes wird getrennt; Benutzer wird abgemeldet
225 Data connection open; no transfer in progress 					Datenverbindung hergestellt; derzeit keine Übertragung
226 Closing data connection. Requested file action successful 		Datenverbindung wird getrennt
227 Entering Passive Mode 										Passiver Modus aktiviert
230 User logged in, proceed 									Benutzer angemeldet, bitte fortfahren
250 Requested file action okay, completed 						Angeforderter Vorgang OK, beendet
257 "PATH" created 											"PFAD" wurde erstellt
331 User name okay, need password 							Benutzername OK, Kennwort erforderlich
332 Need account for login 										Benutzerkonto zur Anmeldung erforderlich
350 Requested file action pending further information 				Mehr Informationen für Dateivorgang erforderlich
421 Service not available, closing control connection 				Dienst nicht verfügbar, Steuerverbindung wird getrennt
425 Can't open data connection 									Datenverbindung kann nicht hergestellt werden
426 Connection closed; transfer aborted Verbindung getrennt; 		Übertragung abgebrochen
450 Requested file action not taken; File unavailable 				Angeforderter Dateivorgang wurde nicht ausgeführt; Datei nicht verfügbar
451 Requested action aborted: local error in processing 				Angeforderter Vorgang abgebrochen: Lokaler Fehler bei der Bearbeitung
452 Requested action not taken; Insufficient storage space in system 	Angeforderter Vorgang nicht ausgeführt; Nicht genügend Speicherplatz auf System
500 Syntax error 												Befehl nicht erkannt
501 Syntax error in parameters or arguments 						Syntaxfehler bei den Parametern
502 Command not implemented 									Befehl nicht implementiert
503 Bad sequence of commands 								Ungültige Befehlsabfolge
504 Command not implemented for that parameter 					Befehl für diesen Parameter nicht implementiert
530 Not logged in 												Nicht angemeldet
532 Need account for storing files 								Zum Speichern von Dateien Anmeldung erforderlich
550 Requested file action not taken; File unavailable Angeforderter 	Dateivorgang wurde nicht ausgeführt; Datei nicht verfügbar
551 Requested action aborted: page type unknown 					Angeforderter Vorgang abgebrochen: Unbekannter Seitentyp
552 Requested file action aborted: Exceeded storage allocation 		Angeforderter Dateivorgang abgebrochen: Nicht genügend Platz in aktuellem Verzeichnis oder Datensatz
553 Requested action not taken: File name not allowed 				Angeforderter Vorgang nicht ausgeführt: Unzulässiger Dateiname

#########################
ERROR_T

1 = DNS_CLIENT
2 = FTP Steuerkanal
3 = FTP Datenkanal
4 = FILE_SERVER
5 = Ablaufstörung
#########################

*)

(*@KEY@:END_DESCRIPTION*)
FUNCTION_BLOCK FTP_CLIENT

(*Group:debug*)

VAR
	(*<LOG_MSG :	LOG_MSG;>*)(*Debug-Bausteininstanz*)
END_VAR

VAR_EXTERNAL
	(*<LOG_CL :	us_LOG_CONTROL;>*)(*Debug-Datenstruktur*)
END_VAR

VAR
	(*<_debug_enable :	BOOL := TRUE;>*)
END_VAR

(*Group:parameter*)

VAR_INPUT
	ACTIVATE :	BOOL;
	FILENAME :	STRING;
	FTP_URL :	oscat_STRING250;
	FTP_DOWNLOAD :	BOOL;
	FTP_ACTIV :	BOOL;
	FILE_DELETE :	BOOL;
	TIMEOUT :	TIME;
	DNS_IP4 :	DWORD;
	PLC_IP4 :	DWORD;
END_VAR

VAR_OUTPUT
	DONE :	BOOL;
	BUSY :	BOOL;
	ERROR_C :	DWORD;
	ERROR_T :	BYTE;
END_VAR

(*Group:Default*)

VAR
	IP_C1 :	oscat_IP_C;
	IP_C2 :	oscat_IP_C;
	S_BUF1 :	oscat_NETWORK_BUFFER;
	S_BUF2 :	oscat_NETWORK_BUFFER;
	R_BUF1 :	oscat_NETWORK_BUFFER;
	R_BUF2 :	oscat_NETWORK_BUFFER;
	URL_DATA :	oscat_url;
	DNS_CLIENT :	DNS_CLIENT;
	IPC1 :	IP_CONTROL;
	IPC2 :	IP_CONTROL;
	FS :	FILE_SERVER;
	FSD :	oscat_FILE_SERVER_DATA;
	activate_last :	BOOL;
	step :	INT;
	snd_step :	INT;
	snd_text :	oscat_STRING250;
	rcv_text :	oscat_STRING250;
	rcv_state :	INT;
	TON_WAIT :	TON;
	last_step :	INT;
	next_step :	INT;
	idx1 :	INT;
	idx2 :	INT;
	str1 :	oscat_STRING250;
	str2 :	oscat_STRING250;
	ftp_path :	STRING;
	byar :	oscat_aB0_5;
	dw_tmp :	DWORD;
	w_tmp :	WORD;
	fpd :	oscat_FILE_PATH_DATA;
	timeout2 :	TIME;
	timeout3 :	TIME;
	ip_c1_red_disable :	BOOL;(*IP_CONTROL 1 - Remote Disconnect Error unterdrücken*)
	ip_c2_red_disable :	BOOL;(*IP_CONTROL 2 - Remote Disconnect Error unterdrücken*)
	ftp_file_size :	UDINT;
	STRING_TO_URL :	STRING_TO_URL;
	BUFFER_TO_STRING :	BUFFER_TO_STRING_NW;
	_STRING_TO_BUFFER :	_STRING_TO_BUFFER_NW;
	ELEMENT_GET :	ELEMENT_GET;
	FILE_PATH_SPLIT :	FILE_PATH_SPLIT;
	IS_NUM :	IS_NUM;
END_VAR

(*@KEY@: WORKSHEET
NAME: FTP_CLIENT
IEC_LANGUAGE: ST
*)

CASE step OF

00:	IF ACTIVATE AND NOT activate_last THEN
		ftp_file_size := UDINT#0;
		TIMEOUT := MAX(T#10s,TIMEOUT);
		timeout2 := TIMEOUT + T#1s;
		timeout3 := DIV_T_AI(TIMEOUT,2);
		DONE := FALSE;
		ip_c1_red_disable := FALSE;
		ip_c2_red_disable := FALSE;
		ERROR_C := DWORD#0;
		ERROR_T := BYTE#0;
		FSD.ERROR := BYTE#0;
		STRING_TO_URL(STR:=FTP_URL,DEFAULT_PROTOCOL:='',DEFAULT_PATH:='/');
		URL_DATA := STRING_TO_URL.STRING_TO_URL;
		IF LEN(URL_DATA.USER) = 0 THEN
			URL_DATA.USER := 'Anonymous';
			URL_DATA.PASSWORD := 'User@';
		END_IF;

		FILE_PATH_SPLIT(FILENAME:=FILENAME,X:=fpd); (* Datei-Path zerlegen *)
		fpd := FILE_PATH_SPLIT.X;
		str1 := fpd.FILENAME; (* zwischenspeichern *)
		FILE_PATH_SPLIT(FILENAME:=URL_DATA.PATH,X:=fpd); (* FTP-Path zerlegen *)
		fpd := FILE_PATH_SPLIT.X;
		IF LEN(fpd.FILENAME) = 0 THEN (* wenn FTP-Path keinen Dateinamen enthält , dann den Namen der lokalen Datei benutzen *)
			ftp_path := CONCAT(URL_DATA.PATH,str1);
		ELSE
			ftp_path := URL_DATA.PATH;
		END_IF;
		step := 10;
	END_IF;

10:	IF DNS_CLIENT.DONE THEN
		step := 20;
	ELSIF DNS_CLIENT.ERROR <> DWORD#0 THEN
		ERROR_C := DNS_CLIENT.ERROR;
		ERROR_T := BYTE#1;
		step := 980;
	END_IF;

20:	(* FTP Steuerkanal einrichten *)
	IP_C1.C_PORT := WORD#21; (* Portnummer eintragen *)
  	IP_C1.C_IP := DNS_CLIENT.IP4; (* IP eintragen *)
  	IP_C1.C_MODE := BYTE#0; (* Mode: TCP+ACTIV+PORT *)
  	IP_C1.TIME_RESET := TRUE; (* Zeitueberwachung rücksetzen *)
  	IP_C1.C_ENABLE := TRUE; (* Verbindungsaufbau freigeben *)
  	IP_C1.R_OBSERVE := TRUE; (* Empfangsueberwachung *)
	R_BUF1.SIZE := UINT#0;

  	IP_C2.C_ENABLE   := FALSE; (* Verbindungsaufbau sperren *)
	step := 30;

30:	IF rcv_state = 220 THEN (* 220 = Service ready for new user *)
		snd_text := CONCAT('USER ',URL_DATA.USER);
		next_step := 40;
	END_IF;

40:	IF rcv_state = 331 THEN (* 331 = User name okay, need password *)
		snd_text := CONCAT('PASS ',URL_DATA.PASSWORD);
		next_step := 50;
	ELSIF rcv_state = 230 THEN (* 230 = User logged in, proceed *)
		next_step := 50;
	ELSIF rcv_state = 220 THEN (* 220 = Service ready for new user *)
		next_step := 20; (* WORK verbindung sollte ab/aufgebaut werden *)
	END_IF;

50:	IF rcv_state = 230 THEN (* 230 = User logged in, proceed *)
		snd_text := 'TYPE I';  (* binären Modus aktivieren *)
		next_step := 54;
	END_IF;

54:	IF rcv_state = 200 THEN (* 200 = Command okay *)
		IF FTP_DOWNLOAD THEN (* Datei von FTP Empfangen *)
			snd_text := CONCAT('SIZE ', ftp_path); (* SIZE /PFAD/FILENAME *)
			next_step := 56;
		ELSE
			step := 60;
		END_IF;
	END_IF;

56:	IF rcv_state = 213 THEN (* 213 Filesize *)
		ELEMENT_GET(SEP:=BYTE#32,POS:=1,ELEMENT:=rcv_text);
		rcv_text := ELEMENT_GET.ELEMENT;
		str1 := ELEMENT_GET.ELEMENT_GET;
		ftp_file_size := STRING_TO_UDINT(str1); (* Dateigroesse in bytes gestimmen *)
		step := 60;
	END_IF;

60:	IF FTP_ACTIV THEN (* FTP Server aktiv *)
		IF URL_DATA.PORT = WORD#0 THEN
			URL_DATA.PORT := WORD#20; (* Standard Datenkanal *)
		END_IF;
		str2 := '';
		dw_tmp := PLC_IP4;
		FOR idx1 := 0 TO 5 DO
			IF idx1 = 4 THEN
				dw_tmp := ROR(WORD_TO_DWORD(URL_DATA.PORT),8);
			ELSE
				dw_tmp := ROL(dw_tmp,8);
			END_IF;
			str2 := CONCAT(str2,BYTE_TO_STRING(DWORD_TO_BYTE(dw_tmp),'%u'));
			IF idx1 < 5 THEN
				str2 := CONCAT(str2,',');
			END_IF;
		END_FOR;
		dw_tmp := DNS_CLIENT.IP4; (* IP eintragen *)
		w_tmp := URL_DATA.PORT; (* Port Nummer des Datenkanals *)
		snd_text := CONCAT('PORT ',str2); (* FTP Server in den aktiv-mode schalten *)
		next_step := 80;
	ELSE
		snd_text := 'PASV';  (* FTP Server in den passiv-mode schalten *)
		next_step := 70;
	END_IF;
	step := 999; (* Warten auf next_step *)

70:	IF rcv_state = 227 THEN (* 227 = Entered Passive Mode (213,202,225,43,212,186) *)
		idx1 := FIND(rcv_text , '(' );
		idx2 := FIND(rcv_text , ')' );
		IF idx1 > 0 AND idx2 > idx1+1 THEN
			str1 := MID(rcv_text, idx2 - idx1 - 1, idx1+1);
			FOR idx1 := 0 TO 5 DO
				ELEMENT_GET(SEP:=BYTE#44,POS:=idx1,ELEMENT:=str1);
				str1 := ELEMENT_GET.ELEMENT;
				str2 := ELEMENT_GET.ELEMENT_GET;
				byar[idx1] := STRING_TO_BYTE(str2);
			END_FOR;
			dw_tmp := DWORD_OF_BYTE(byar[0],byar[1],byar[2],byar[3]); (* IP Adresse des Datenkanals *)
			w_tmp := WORD_OF_BYTE(byar[4],byar[5]); (* Port Nummer des Datenkanals *)
		END_IF;
		step := 100;
	END_IF;

80:	IF rcv_state = 200 THEN (* 200 = PORT command successful *)
		step := 100;
	END_IF;

100:IP_C2.C_MODE := SEL(FTP_ACTIV,BYTE#0,BYTE#2); (* Aktiv = Mode 2: TCP+PASSIV+PORT / passiv = Mode 0: TCP+ACTIV+PORT *)
	IP_C2.C_IP := dw_tmp; (* IP Adresse des Datenkanals *)
	IP_C2.C_PORT := w_tmp; (* Port Nummer des Datenkanals *)
  	IP_C2.TIME_RESET := TRUE; (* Zeitueberwachung rücksetzen *)
  	IP_C2.C_ENABLE := TRUE; (* Verbindungsaufbau freigeben *)
	IP_C2.R_OBSERVE := FALSE; (* Empfangsueberwachung *)
	R_BUF2.SIZE := UINT#0;
	step := 120;

120:IF IP_C2.C_STATE > BYTE#127 THEN (* FTP Datenkanal aufgebaut *)
		IF FTP_DOWNLOAD THEN (* File von FTP empfangen *)
			IP_C2.MAILBOX[3] := BYTE#1; (* IP Empfang sperren *)
			step := 400;
		ELSE
			snd_text := 'STOR ';
			next_step := 140;
			snd_text := CONCAT(snd_text, ftp_path); (* STORE /PFAD/FILENAME *)
			step := 999; (* Warten auf next_step *)
		END_IF;
	END_IF;

(* ============== File an FTP senden ================ *)

140:IF rcv_state = 125 OR rcv_state = 150 THEN (* 125 = Data connection already open / 150 = File status okay; about to open data connection *)
		step := 160;
	END_IF;

160:FSD.FILENAME := FILENAME; (* Dateiname *)
	FSD.MODE := BYTE#1; (* vorhandene Datei zum lesen öffnen *)
	FSD.OFFSET := UDINT#0; (* Start bei Dateianfang *)
	FSD.AUTO_CLOSE := T#0s; (* kein Auto-Close verwenden *)
	S_BUF2.SIZE := UINT#65535; (* maximale länge einlesen *)
	IP_C2.MAILBOX[2] := BYTE#1; (* IP Senden blockieren *)
	step := 200;

200:IF FSD.MODE = BYTE#0 AND FSD.ERROR = BYTE#0 THEN
		IP_C2.MAILBOX[2] := BYTE#0; (* IP Senden erlauben *)
		step := 210;
	END_IF;

210:IF S_BUF2.SIZE = UINT#0 THEN (* warten bis alle daten gesendet sind *)
		IF FSD.FILE_SIZE - FSD.OFFSET > UDINT#0 THEN
			FSD.MODE := BYTE#1; (* vorhandene Datei zum lesen öffnen *)
			S_BUF2.SIZE := UINT#65535; (* maximale länge einlesen *)
			IP_C2.MAILBOX[2] := BYTE#1; (* IP Senden blockieren *)
			step := 200;
		ELSE
			IP_C2.C_ENABLE := FALSE; (* FTP Datenkanal schliessen *)
			step := 300;
		END_IF;
	END_IF;

300:IF rcv_state = 226 THEN (* 226 Closing data connection. Requested file action successful  *)
		snd_text := 'QUIT';
		ip_c1_red_disable := TRUE;
		next_step := 320;
	END_IF;

320:IF rcv_state = 221 OR TON_WAIT.ET > timeout3  THEN (* 221 Service closing control connection *)
		IP_C1.C_ENABLE := FALSE; (* FTP Steuerkanal schliessen *)
		IF FILE_DELETE THEN (* Datei nach transfer löschen *)
			FSD.MODE := BYTE#4; (* File Remove *)
			step := 340;
		ELSE
			step := 900;
		END_IF;
	END_IF;

340:IF FSD.MODE = BYTE#0 AND FSD.ERROR = BYTE#0 THEN
		step := 900;
	END_IF;

(*  ============== File vom FTP Empfangen  ============== *)

400:snd_text := 'RETR ';
	next_step := 410;
	snd_text := CONCAT(snd_text, ftp_path); (* RETR /PFAD/FILENAME *)
	step := 999; (* Warten auf next_step *)

410:IF rcv_state = 125 OR rcv_state = 150 THEN (* 125 = Data connection already open / 150 = File status okay; about to open data connection *)
		IP_C2.R_OBSERVE := TRUE; (* Empfangsueberwachung *)
		step := 420;
	END_IF;

420:FSD.FILENAME := FILENAME; (* Dateiname *)
	FSD.MODE := BYTE#3; (* Datei neu anlegen *)
	FSD.OFFSET := UDINT#0; (* Start bei Dateianfang *)
	FSD.AUTO_CLOSE := T#0s; (* kein Auto-Close verwenden *)
	step := 460;

440:IF R_BUF2.SIZE > UINT#0 THEN (* warten bis daten empfangen wurden *)
		IP_C2.MAILBOX[3] := BYTE#1; (* IP Empfang blockieren bis Daten in Datei geschrieben wurden *)
		FSD.MODE := BYTE#3; (* Daten in Datei schreiben *)
		step := 460;
	ELSIF FSD.FILE_SIZE = ftp_file_size THEN (* Verbindung abgebaut ? , oder 226 = Closing data connection. Requested file action successful *)
		IP_C2.C_ENABLE := FALSE; (* FTP Datenkanal schliessen *)
		ip_c2_red_disable := TRUE;
		step := 700;
	END_IF;

460:IF FSD.MODE = BYTE#0 AND FSD.ERROR = BYTE#0 THEN (* warten bis Daten geschreiben wurden *)
		R_BUF2.SIZE := UINT#0; (* Daten löschen *)
		IP_C2.MAILBOX[3] := BYTE#0; (* IP Empfang wieder erlauben *)
		step := 440;
	END_IF;

(* ================================================== *)

700:IF rcv_state = 226 OR  TON_WAIT.ET > timeout3 THEN (* 226 Closing control connection. Requested file action successful  *)
		IF FTP_DOWNLOAD AND FILE_DELETE THEN (* FTP Download und File löschen ? *)
			snd_text := CONCAT('DELE ', ftp_path); (* DELE /PFAD/FILENAME *)
			next_step := 720;
		ELSE
			step := 740;
		END_IF;
	END_IF;

720:IF rcv_state = 250 THEN (* 250 Requested file action okay, completed *)
		step := 740;
	END_IF;

740:snd_text := 'QUIT';
	ip_c1_red_disable := TRUE;
	next_step := 760;
	step := 999; (* Warten auf next_step *)

760:IF rcv_state = 221 OR TON_WAIT.ET > timeout3 THEN (* 221 Service closing control connection  *)
		IP_C1.C_ENABLE := FALSE; (* FTP Steuerkanal schliessen *)
		IF NOT FTP_DOWNLOAD AND FILE_DELETE THEN (* FTP Upload und Datei nach transfer löschen *)
			FSD.MODE := BYTE#4; (* File Remove *)
			step := 780;
		ELSE
			step := 900;
		END_IF;
	END_IF;

780:IF FSD.MODE = BYTE#0 AND FSD.ERROR = BYTE#0 THEN
		step := 900;
	END_IF;

(* ================================================== *)

900:DONE := TRUE;
	step := 980;

980:IP_C1.C_ENABLE := FALSE; (* FTP Steuerkanal schliessen *)
	IP_C2.C_ENABLE := FALSE; (* FTP Datenkanal schliessen *)
	IP_C2.MAILBOX[2] := BYTE#0; (* IP Senden wieder erlauben *)
	IP_C2.MAILBOX[3] := BYTE#0; (* IP Empfang wieder erlauben *)
	S_BUF1.SIZE := UINT#0;
	S_BUF2.SIZE := UINT#0;
	R_BUF1.SIZE := UINT#0;
	R_BUF2.SIZE := UINT#0;
	ftp_file_size := UDINT#0;
	snd_step := 0;
	next_step := 0;
	FSD.MODE := BYTE#5; (* Datei schliessen *)
	step := 990;

990:IF IP_C1.C_STATE = BYTE#0 AND IP_C2.C_STATE = BYTE#0 AND FSD.FILE_OPEN = FALSE THEN
		step := 0;
	END_IF;

999: ; (* Dummy Schritt, warten bis neuer schritt durch "next_step" aktiv wird *)

END_CASE;

(* ++++++++++++++++++++++++++++++++++++++++++++++++++++++++++ *)

IF step >= 30 THEN
	IF R_BUF1.SIZE > UINT#0 THEN (* Daten wurden empfangen ? *)
		idx1 := UINT_TO_INT(R_BUF1.SIZE);
		REPEAT (* zeilenterminierung erkennen und echtes TEXT-Ende bestimmen *)
			idx1 := idx1 - 1;
		UNTIL idx1 = 0 OR R_BUF1.BUFFER[idx1] >= BYTE#32 (* TRUE = EXIT *)
		END_REPEAT;
		idx1 := idx1 + 1; (* index auf SIZE umrechnen *)
		BUFFER_TO_STRING(PT:=R_BUF1.BUFFER,SIZE:=INT_TO_UINT(idx1),START:=UINT#0,STOP:=UINT#249);
		R_BUF1.BUFFER := BUFFER_TO_STRING.PT;
		rcv_text := BUFFER_TO_STRING.BUFFER_TO_STRING;
		IF LEN(rcv_text) >= 3 THEN (* Statuscode prüfen und auswerten *)
			str1 := LEFT(rcv_text,3);
			IS_NUM(STR:=str1);
			IF IS_NUM.IS_NUM THEN (* enthält nur Zahlen ? *)
				rcv_state := STRING_TO_INT(str1);
			END_IF;
			IP_C1.R_OBSERVE := FALSE;
		END_IF;
		R_BUF1.SIZE := UINT#0; (* daten löschen *)

        (*####################  DEBUG-MESSAGE  ###################################*)
        (*IF _debug_enable THEN
          LOG_CL.NEW_MSG := '(~D ~T) RCV: >~1<';
          LOG_CL.PRINTF[1] := rcv_text;
          LOG_MSG();
        END_IF;*)
        (*########################################################################*)

	END_IF;
END_IF;

(* automatisches Datensenden *)

CASE snd_step OF

00:	IF LEN(snd_text) > 0 THEN

        (*####################  DEBUG-MESSAGE  ###################################*)
        (*IF _debug_enable THEN
          LOG_CL.NEW_MSG := '(~D ~T) SND: >~1<';
          LOG_CL.PRINTF[1] := snd_text;
          LOG_MSG();
        END_IF;*)
        (*########################################################################*)

		_STRING_TO_BUFFER(STR:=snd_text,POS:=0,SIZE:=UINT#4096,PT:=S_BUF1.BUFFER); (* String in puffer kopieren *)
		S_BUF1.BUFFER := _STRING_TO_BUFFER.PT;
		idx1 := LEN(snd_text);
		S_BUF1.BUFFER[idx1] := BYTE#16#0D;
		idx1 := idx1 + 1;
		S_BUF1.BUFFER[idx1] := BYTE#16#0A;
		idx1 := idx1 + 1;
		S_BUF1.SIZE := INT_TO_UINT(idx1); (* Sendelänge eintragen *)
		R_BUF1.SIZE := UINT#0; (* Empfangsbuffer rücksetzen *)
		IP_C1.R_OBSERVE := TRUE;
		rcv_state := 9999; (* letzen FTP Status löschen *)
		snd_text := '';
		snd_step := 10;

	END_IF;

10:	IF S_BUF1.SIZE = UINT#0 THEN (* warten bis alle daten gesendet sind *)
		step := next_step;
		snd_step := 0;
	END_IF;

END_CASE;

(* Globale Fehlerbehandlung für Haupt-Routine *)
IF ERROR_T = BYTE#0 AND step > 20 THEN (* noch kein Fehler gespeichert und Hauptroutine aktiv *)

	IF IP_C1.ERROR > DWORD#0 AND IP_C1.C_ENABLE AND NOT IP_C1.TIME_RESET THEN  (* IP Control 1 *)
		IF ip_c1_red_disable = FALSE OR IP_C1.ERROR <> DWORD#16#FD000000 THEN
			ERROR_C := IP_C1.ERROR;
			ERROR_T := BYTE#2;
			step := 980;
		END_IF;
	END_IF;

	IF IP_C2.ERROR > DWORD#0 AND IP_C2.C_ENABLE AND NOT IP_C2.TIME_RESET THEN  (* IP Control 2 *)
		IF ip_c2_red_disable = FALSE OR IP_C2.ERROR <> DWORD#16#FD000000 THEN
			ERROR_C := IP_C2.ERROR;
			ERROR_T := BYTE#3;
			step := 980;
		END_IF;
	END_IF;

	IF FSD.MODE = BYTE#0 THEN
		IF FSD.ERROR > BYTE#0 THEN
			ERROR_C := BYTE_TO_DWORD(FSD.ERROR);
			ERROR_T := BYTE#4; (* Dateizugriff *)
			step := 980;
		END_IF;
	END_IF;
END_IF;

IF TON_WAIT.Q THEN (* Ablaufstörung - Schrittkette *)
	ERROR_C := SHL(INT_TO_DWORD(step),16) OR INT_TO_DWORD(rcv_state); (* aktuellen Schritt und letzten FTP Status eintragen *)
	ERROR_T := BYTE#5;
	step := 980;
END_IF;

(* ######################################################## *)

DNS_CLIENT(IP_C:=IP_C1, S_BUF:=S_BUF1, R_BUF:=R_BUF1, DOMAIN:=URL_DATA.DOMAIN, IP4_DNS:= DNS_IP4, ACTIVATE:=step=10); (* DNS-Client *)
IP_C1  := DNS_CLIENT.IP_C;
R_BUF1 := DNS_CLIENT.R_BUF;
S_BUF1 := DNS_CLIENT.S_BUF;

IPC1(IP:= DWORD#0, PORT:= WORD#0 , TIME_OUT:= TIMEOUT, IP_C:= IP_C1, S_BUF:= S_BUF1, R_BUF:= R_BUF1); (* FTP Steuerkanal *)
IP_C1  := IPC1.IP_C;
R_BUF1 := IPC1.R_BUF;
S_BUF1 := IPC1.S_BUF;

IPC2(IP:= DWORD#0, PORT:= WORD#0 , TIME_OUT:= TIMEOUT, IP_C:= IP_C2, S_BUF:= S_BUF2, R_BUF:= R_BUF2); (* FTP Datenkanal *)
IP_C2  := IPC2.IP_C;
R_BUF2 := IPC2.R_BUF;
S_BUF2 := IPC2.S_BUF;

TON_WAIT(IN:=step = last_step AND step > 0,PT:=timeout2);
last_step := step;
activate_last := ACTIVATE;
BUSY := step <> 0;

IF FTP_DOWNLOAD THEN (* FILE_SERVER *)
	FS(FSD:=FSD,PT:=R_BUF2); (* Datei von FTP empfangen *)
	FSD    := FS.FSD;
	R_BUF2 := FS.PT;
ELSE
	FS(FSD:=FSD,PT:=S_BUF2); (* Datei an FTP senden *)
	FSD	   := FS.FSD;
	S_BUF2 := FS.PT;
END_IF;

(* revision history
ks	11. may 2011	rev 1.2
	ip_control - remote disconnect error ausblenden, und sonderbehandlung für pcworx

ks	06. apr. 2011	rev 1.1
	list_len und list_get durch element_count und element_get ersetzt

ks	01. jan. 2011	rev 1.0
	original version
*)

(*@KEY@: END_WORKSHEET *)
END_FUNCTION_BLOCK
